   #FRK_JsonHeader := FALSE;
   #Line := WSTRING#'{';
   #Ok := "FRK_JsonAdd"(Key := 'set', Value := STRING_TO_WSTRING(#Data.SetName), Quoted := TRUE, LastField := FALSE, Line := #Line);
   IF NOT #Ok THEN
       #Line := WSTRING#'';
       RETURN;
   END_IF;
   #Ok := "FRK_JsonAdd"(Key := 'root', Value := STRING_TO_WSTRING(#Data.RootIdentity), Quoted := TRUE, LastField := FALSE, Line := #Line);
   IF NOT #Ok THEN
       #Line := WSTRING#'';
       RETURN;
   END_IF;
   #Ok := "FRK_JsonAdd"(Key := 'schema', Value := UINT_TO_WSTRING(#Data.SetSchema), Quoted := FALSE, LastField := FALSE, Line := #Line);
   IF NOT #Ok THEN
       #Line := WSTRING#'';
       RETURN;
   END_IF;
   #Ok := "FRK_JsonAdd"(Key := 'configRev', Value := UDINT_TO_WSTRING(#Data.ConfigRev), Quoted := FALSE, LastField := FALSE, Line := #Line);
   IF NOT #Ok THEN
       #Line := WSTRING#'';
       RETURN;
   END_IF;
   #Ok := "FRK_JsonAdd"(Key := 'kind', Value := DINT_TO_WSTRING(#Data.Kind), Quoted := FALSE, LastField := FALSE, Line := #Line);
   IF NOT #Ok THEN
       #Line := WSTRING#'';
       RETURN;
   END_IF;
   #Ok := "FRK_JsonAdd"(Key := 'model', Value := STRING_TO_WSTRING(#Data.ModelCode), Quoted := TRUE, LastField := FALSE, Line := #Line);
   IF NOT #Ok THEN
       #Line := WSTRING#'';
       RETURN;
   END_IF;
   #Ok := "FRK_JsonAdd"(Key := 'records', Value := DINT_TO_WSTRING(#Data.RecordCount), Quoted := FALSE, LastField := FALSE, Line := #Line);
   IF NOT #Ok THEN
       #Line := WSTRING#'';
       RETURN;
   END_IF;
   #Ok := "FRK_JsonAdd"(Key := 'created', Value := ULINT_TO_WSTRING(LDT_TO_ULINT(#Data.CreatedAt) / ULINT#1000000000), Quoted := FALSE, LastField := FALSE, Line := #Line);
   IF NOT #Ok THEN
       #Line := WSTRING#'';
       RETURN;
   END_IF;
   IF #Data.TimeSynchronized THEN
       #Flag := WSTRING#'1';
   ELSE
       #Flag := WSTRING#'0';
   END_IF;
   #Ok := "FRK_JsonAdd"(Key := 'clock', Value := #Flag, Quoted := FALSE, LastField := TRUE, Line := #Line);
   IF NOT #Ok THEN
       #Line := WSTRING#'';
       RETURN;
   END_IF;
   #FRK_JsonHeader := TRUE;
END_FUNCTION

FUNCTION "FRK_JsonParse" : Bool   // FC110, SCL
{ S7_Optimized_Access := 'TRUE' }
VERSION : 0.1
// Strict flat JSON object scanner: whole object, unique known fields, exact
//  types, numeric integer grammar; strings decode escapes before owner checks.
// stored: AutoNumber true, IsIECCheckEnabled false, SetENOAutomatically false, UDAEnableTagReadback false
   VAR_INPUT
      Line : WString;
   END_VAR
   VAR_IN_OUT
      Fields : Array[1..9] of "FRK_JsonField";
      Count : Int;
   END_VAR
   VAR_TEMP
      Pos : Int;
      Limit : Int;
      Digit : Int;
      CodePoint : UInt;
      HexIndex : Int;
      Index : Int;
      Part : Int;
      Text : WString[160];
      Piece : WString[1];
      Quoted : Bool;
      Closed : Bool;
      Ch : WChar;
   END_VAR
BEGIN

   #FRK_JsonParse := FALSE;
   #Count := 0;
   #Pos := 1;
   #Limit := LEN(#Line);
   IF #Limit < 2 OR #Line[#Pos] <> WCHAR#'{' THEN
       RETURN;
   END_IF;
   #Pos := #Pos + 1;
   WHILE #Pos <= #Limit DO
       "FRK_JsonSkip"(Line := #Line,
                      Pos := #Pos);
       IF #Pos > #Limit OR #Count >= 9 THEN
           RETURN;
       END_IF;
       #Count := #Count + 1;
       FOR #Part := 1 TO 2 DO
           #Text := WSTRING#'';
           #Closed := FALSE;
           #Quoted := #Line[#Pos] = WCHAR#'"';
           IF #Part = 1 AND NOT #Quoted THEN
               RETURN;
           END_IF;
           IF #Quoted THEN
               #Pos := #Pos + 1;
           END_IF;
           WHILE #Pos <= #Limit DO
               #Ch := #Line[#Pos];
               IF #Quoted AND #Ch = WCHAR#'"' THEN
                   #Closed := TRUE;
                   #Pos := #Pos + 1;
                   EXIT;
               END_IF;
               IF NOT #Quoted AND (#Ch = WCHAR#',' OR #Ch = WCHAR#'}' OR #Ch = WCHAR#' ') THEN
                   #Closed := TRUE;
                   EXIT;
               END_IF;
               IF #Ch < WCHAR#'$0020' THEN
                   RETURN;
               END_IF;
               IF #Quoted AND #Ch = WCHAR#'\' THEN
                   #Pos := #Pos + 1;
                   IF #Pos > #Limit THEN
                       RETURN;
                   END_IF;
                   #Ch := #Line[#Pos];
                   IF #Ch = WCHAR#'u' THEN
                       #CodePoint := 0;
                       FOR #HexIndex := 1 TO 4 DO
                           #Pos := #Pos + 1;
                           IF #Pos > #Limit THEN
                               RETURN;
                           END_IF;
                           #Ch := #Line[#Pos];
                           #Digit := -1;
                           IF #Ch >= WCHAR#'0' AND #Ch <= WCHAR#'9' THEN
                               #Digit := WORD_TO_INT(WCHAR_TO_WORD(#Ch)) - 48;
                           ELSIF #Ch >= WCHAR#'a' AND #Ch <= WCHAR#'f' THEN
                               #Digit := WORD_TO_INT(WCHAR_TO_WORD(#Ch)) - 87;
                           ELSIF #Ch >= WCHAR#'A' AND #Ch <= WCHAR#'F' THEN
                               #Digit := WORD_TO_INT(WCHAR_TO_WORD(#Ch)) - 55;
                           END_IF;
                           IF #Digit < 0 THEN
                               RETURN;
                           END_IF;
                           #CodePoint := #CodePoint * 16 + INT_TO_UINT(#Digit);
                       END_FOR;
                       IF #CodePoint = 0 OR #CodePoint >= UINT#16#D000 THEN
                           RETURN;
                       END_IF;
                       #Ch := WORD_TO_WCHAR(UINT_TO_WORD(#CodePoint));
                   ELSIF #Ch = WCHAR#'n' THEN
                       #Ch := WCHAR#'$000A';
                   ELSIF #Ch = WCHAR#'r' THEN
                       #Ch := WCHAR#'$000D';
                   ELSIF #Ch = WCHAR#'t' THEN
                       #Ch := WCHAR#'$0009';
                   ELSIF #Ch = WCHAR#'b' THEN
                       #Ch := WCHAR#'$0008';
                   ELSIF #Ch = WCHAR#'f' THEN
                       #Ch := WCHAR#'$000C';
                   ELSIF #Ch <> WCHAR#'"' AND #Ch <> WCHAR#'\' AND #Ch <> WCHAR#'/' THEN
                       RETURN;
                   END_IF;
               ELSIF NOT #Quoted AND (#Ch < WCHAR#'0' OR #Ch > WCHAR#'9') THEN
                   RETURN;
               END_IF;
               IF LEN(#Text) >= 160 THEN
                   RETURN;
               END_IF;
               #Piece := WSTRING#' ';
               #Piece[1] := #Ch;
               #Text := CONCAT(IN1 := #Text, IN2 := #Piece);
               #Pos := #Pos + 1;
           END_WHILE;
           IF NOT #Closed THEN
               RETURN;
           END_IF;
           IF #Part = 1 THEN
               IF LEN(#Text) < 1 OR LEN(#Text) > 16 THEN
                   RETURN;
               END_IF;
               #Fields[#Count].Key := WSTRING_TO_STRING(#Text);
               FOR #Index := 1 TO #Count - 1 DO
                   IF #Fields[#Index].Key = #Fields[#Count].Key THEN
                       RETURN;
                   END_IF;
               END_FOR;
               "FRK_JsonSkip"(Line := #Line,
                              Pos := #Pos);
               IF #Pos > #Limit THEN
                   RETURN;
               END_IF;
               IF #Line[#Pos] <> WCHAR#':' THEN
                   RETURN;
               END_IF;
               #Pos := #Pos + 1;
               "FRK_JsonSkip"(Line := #Line,
                              Pos := #Pos);
               IF #Pos > #Limit THEN
                   RETURN;
               END_IF;
           ELSE
               IF NOT #Quoted AND (LEN(#Text) = 0 OR (LEN(#Text) > 1 AND #Text[1] = WCHAR#'0')) THEN
                   RETURN;
               END_IF;
               #Fields[#Count].Text := #Text;
               #Fields[#Count].Quoted := #Quoted;
           END_IF;
       END_FOR;
       "FRK_JsonSkip"(Line := #Line,
                      Pos := #Pos);
       IF #Pos > #Limit THEN
           RETURN;
       END_IF;
       IF #Line[#Pos] = WCHAR#'}' THEN
           #Pos := #Pos + 1;
           "FRK_JsonSkip"(Line := #Line,
                          Pos := #Pos);
           #FRK_JsonParse := #Pos > #Limit;
           RETURN;
       END_IF;
       IF #Line[#Pos] <> WCHAR#',' THEN
           RETURN;
       END_IF;
       #Pos := #Pos + 1;
   END_WHILE;
END_FUNCTION

FUNCTION "FRK_JsonPut" : Bool   // FC108, SCL
{ S7_Optimized_Access := 'TRUE' }
VERSION : 0.1
// Append complete text or refuse. Explicit destination width and length check
//  protect long WSTRING lines against truncation in the Siemens string runtime.
// stored: AutoNumber true, IsIECCheckEnabled false, SetENOAutomatically false, UDAEnableTagReadback false
   VAR_INPUT
      Text : WString;
   END_VAR
   VAR_IN_OUT
      Line : WString;
   END_VAR
   VAR_TEMP
      Expected : Int;
   END_VAR
BEGIN

   #FRK_JsonPut := FALSE;
   #Expected := LEN(#Line) + LEN(#Text);
   IF #Expected > 480 THEN
       RETURN;
   END_IF;
   #Line := CONCAT(IN1 := #Line, IN2 := #Text);
   #FRK_JsonPut := LEN(#Line) = #Expected;
END_FUNCTION

FUNCTION "FRK_JsonReadHeader" : Bool   // FC119, SCL
{ S7_Optimized_Access := 'TRUE' }
VERSION : 0.1
// stored: AutoNumber true, IsIECCheckEnabled false, SetENOAutomatically false, UDAEnableTagReadback false
   VAR_INPUT
      Count : Int;
      Fields : Array[1..9] of "FRK_JsonField";
   END_VAR
   VAR_IN_OUT
      Data : "ST_ConfigSetInfo";
   END_VAR
   VAR_TEMP
      Candidate : "ST_ConfigSetInfo";
      Index : Int;
      Found : Int;
      Ok : Bool;
   END_VAR
BEGIN

   #FRK_JsonReadHeader := FALSE;
   IF #Count <> 9 THEN
       RETURN;
   END_IF;
   #Found := 0;
   FOR #Index := 1 TO #Count DO
       IF #Fields[#Index].Key = 'set' THEN
           #Found := #Index;
       END_IF;
   END_FOR;
   IF #Found = 0 THEN
       RETURN;
   END_IF;
   IF #Fields[#Found].Quoted <> TRUE THEN
       RETURN;
   END_IF;
   IF LEN(#Fields[#Found].Text) > 80 OR STRING_TO_WSTRING(WSTRING_TO_STRING(#Fields[#Found].Text)) <> #Fields[#Found].Text THEN
       RETURN;
   END_IF;
   #Candidate.SetName := WSTRING_TO_STRING(#Fields[#Found].Text);
   #Found := 0;
   FOR #Index := 1 TO #Count DO
       IF #Fields[#Index].Key = 'root' THEN
           #Found := #Index;
       END_IF;
   END_FOR;
   IF #Found = 0 THEN
       RETURN;
   END_IF;
   IF #Fields[#Found].Quoted <> TRUE THEN
       RETURN;
   END_IF;
   IF LEN(#Fields[#Found].Text) > 80 OR STRING_TO_WSTRING(WSTRING_TO_STRING(#Fields[#Found].Text)) <> #Fields[#Found].Text THEN
       RETURN;
   END_IF;
   #Candidate.RootIdentity := WSTRING_TO_STRING(#Fields[#Found].Text);
   #Found := 0;
   FOR #Index := 1 TO #Count DO
       IF #Fields[#Index].Key = 'schema' THEN
           #Found := #Index;
       END_IF;
   END_FOR;
   IF #Found = 0 THEN
       RETURN;
   END_IF;
   IF #Fields[#Found].Quoted <> FALSE THEN
       RETURN;
   END_IF;
   #Ok := "FRK_ConfigDecode"(Text := #Fields[#Found].Text, Storage := 4, Minimum := 0.0, Maximum := 65535.0, MaxLength := 0, Value := "FRK_ConfigScratch".Value);
   IF NOT #Ok THEN
       RETURN;
   END_IF;
   #Candidate.SetSchema := LINT_TO_UINT("FRK_ConfigScratch".Value.Number);
   #Found := 0;
   FOR #Index := 1 TO #Count DO
       IF #Fields[#Index].Key = 'configRev' THEN
           #Found := #Index;
       END_IF;
   END_FOR;
   IF #Found = 0 THEN
       RETURN;
   END_IF;
   IF #Fields[#Found].Quoted <> FALSE THEN
       RETURN;
   END_IF;
   #Ok := "FRK_ConfigDecode"(Text := #Fields[#Found].Text, Storage := 4, Minimum := 0.0, Maximum := 4294967295.0, MaxLength := 0, Value := "FRK_ConfigScratch".Value);
   IF NOT #Ok THEN
       RETURN;
   END_IF;
   #Candidate.ConfigRev := LINT_TO_UDINT("FRK_ConfigScratch".Value.Number);
   #Found := 0;
   FOR #Index := 1 TO #Count DO
       IF #Fields[#Index].Key = 'kind' THEN
           #Found := #Index;
       END_IF;
   END_FOR;
   IF #Found = 0 THEN
       RETURN;
   END_IF;
   IF #Fields[#Found].Quoted <> FALSE THEN
       RETURN;
   END_IF;
   #Ok := "FRK_ConfigDecode"(Text := #Fields[#Found].Text, Storage := 4, Minimum := 0.0, Maximum := 1.0, MaxLength := 0, Value := "FRK_ConfigScratch".Value);
   IF NOT #Ok THEN
       RETURN;
   END_IF;
   #Candidate.Kind := LINT_TO_DINT("FRK_ConfigScratch".Value.Number);
   #Found := 0;
   FOR #Index := 1 TO #Count DO
       IF #Fields[#Index].Key = 'model' THEN
           #Found := #Index;
       END_IF;
   END_FOR;
   IF #Found = 0 THEN
       RETURN;
   END_IF;
   IF #Fields[#Found].Quoted <> TRUE THEN
       RETURN;
   END_IF;
   IF LEN(#Fields[#Found].Text) > 64 OR STRING_TO_WSTRING(WSTRING_TO_STRING(#Fields[#Found].Text)) <> #Fields[#Found].Text THEN
       RETURN;
   END_IF;
   #Candidate.ModelCode := WSTRING_TO_STRING(#Fields[#Found].Text);
   #Found := 0;
   FOR #Index := 1 TO #Count DO
       IF #Fields[#Index].Key = 'records' THEN
           #Found := #Index;
       END_IF;
   END_FOR;
   IF #Found = 0 THEN
       RETURN;
   END_IF;
   IF #Fields[#Found].Quoted <> FALSE THEN
       RETURN;
   END_IF;
   #Ok := "FRK_ConfigDecode"(Text := #Fields[#Found].Text, Storage := 4, Minimum := 0.0, Maximum := 3.0, MaxLength := 0, Value := "FRK_ConfigScratch".Value);
   IF NOT #Ok THEN
       RETURN;
   END_IF;
   #Candidate.RecordCount := LINT_TO_INT("FRK_ConfigScratch".Value.Number);
   #Found := 0;
   FOR #Index := 1 TO #Count DO
       IF #Fields[#Index].Key = 'created' THEN
           #Found := #Index;
       END_IF;
   END_FOR;
   IF #Found = 0 THEN
       RETURN;
   END_IF;
   IF #Fields[#Found].Quoted <> FALSE THEN
       RETURN;
   END_IF;
   #Ok := "FRK_ConfigDecode"(Text := #Fields[#Found].Text, Storage := 4, Minimum := 0.0, Maximum := 4294967295.0, MaxLength := 0, Value := "FRK_ConfigScratch".Value);
   IF NOT #Ok THEN
       RETURN;
   END_IF;
   #Candidate.CreatedAt := ULINT_TO_LDT(LINT_TO_ULINT("FRK_ConfigScratch".Value.Number) * ULINT#1000000000);
   #Found := 0;
   FOR #Index := 1 TO #Count DO
       IF #Fields[#Index].Key = 'clock' THEN
           #Found := #Index;
       END_IF;
   END_FOR;
   IF #Found = 0 THEN
       RETURN;
   END_IF;
   IF #Fields[#Found].Quoted <> FALSE THEN
       RETURN;
   END_IF;
   #Ok := "FRK_ConfigDecode"(Text := #Fields[#Found].Text, Storage := 4, Minimum := 0.0, Maximum := 1.0, MaxLength := 0, Value := "FRK_ConfigScratch".Value);
   IF NOT #Ok THEN
       RETURN;
   END_IF;
   #Candidate.TimeSynchronized := "FRK_ConfigScratch".Value.Number = 1;
   #Data := #Candidate;
   #FRK_JsonReadHeader := TRUE;
END_FUNCTION

FUNCTION "FRK_JsonReadRecord" : Bool   // FC121, SCL
{ S7_Optimized_Access := 'TRUE' }
VERSION : 0.1
// stored: AutoNumber true, IsIECCheckEnabled false, SetENOAutomatically false, UDAEnableTagReadback false
   VAR_INPUT
      Count : Int;
      Fields : Array[1..9] of "FRK_JsonField";
   END_VAR
   VAR_IN_OUT
      Data : "ST_ConfigRecord";
   END_VAR
   VAR_TEMP
      Candidate : "ST_ConfigRecord";
      Index : Int;
      Found : Int;
      Ok : Bool;
   END_VAR
BEGIN

   #FRK_JsonReadRecord := FALSE;
   IF #Count <> 6 THEN
       RETURN;
   END_IF;
   #Found := 0;
   FOR #Index := 1 TO #Count DO
       IF #Fields[#Index].Key = 'scope' THEN
           #Found := #Index;
       END_IF;
   END_FOR;
   IF #Found = 0 THEN
       RETURN;
   END_IF;
   IF #Fields[#Found].Quoted <> TRUE THEN
       RETURN;
   END_IF;
   IF LEN(#Fields[#Found].Text) > 80 OR STRING_TO_WSTRING(WSTRING_TO_STRING(#Fields[#Found].Text)) <> #Fields[#Found].Text THEN
       RETURN;
   END_IF;
   #Candidate.Scope := WSTRING_TO_STRING(#Fields[#Found].Text);
   #Found := 0;
   FOR #Index := 1 TO #Count DO
       IF #Fields[#Index].Key = 'key' THEN
           #Found := #Index;
       END_IF;
   END_FOR;
   IF #Found = 0 THEN
       RETURN;
   END_IF;
   IF #Fields[#Found].Quoted <> TRUE THEN
       RETURN;
   END_IF;
   IF LEN(#Fields[#Found].Text) > 160 OR STRING_TO_WSTRING(WSTRING_TO_STRING(#Fields[#Found].Text)) <> #Fields[#Found].Text THEN
       RETURN;
   END_IF;
   #Candidate.WriteKey := WSTRING_TO_STRING(#Fields[#Found].Text);
   #Found := 0;
   FOR #Index := 1 TO #Count DO
       IF #Fields[#Index].Key = 'rev' THEN
           #Found := #Index;
       END_IF;
   END_FOR;
   IF #Found = 0 THEN
       RETURN;
   END_IF;
   IF #Fields[#Found].Quoted <> FALSE THEN
       RETURN;
   END_IF;
   #Ok := "FRK_ConfigDecode"(Text := #Fields[#Found].Text, Storage := 4, Minimum := 0.0, Maximum := 4294967295.0, MaxLength := 0, Value := "FRK_ConfigScratch".Value);
   IF NOT #Ok THEN
       RETURN;
   END_IF;
   #Candidate.Revision := LINT_TO_UDINT("FRK_ConfigScratch".Value.Number);
   #Found := 0;
   FOR #Index := 1 TO #Count DO
       IF #Fields[#Index].Key = 'kind' THEN
           #Found := #Index;
       END_IF;
   END_FOR;
   IF #Found = 0 THEN
       RETURN;
   END_IF;
   IF #Fields[#Found].Quoted <> FALSE THEN
       RETURN;
   END_IF;
   #Ok := "FRK_ConfigDecode"(Text := #Fields[#Found].Text, Storage := 4, Minimum := 0.0, Maximum := 1.0, MaxLength := 0, Value := "FRK_ConfigScratch".Value);
   IF NOT #Ok THEN
       RETURN;
   END_IF;
   #Candidate.Kind := LINT_TO_DINT("FRK_ConfigScratch".Value.Number);
   #Found := 0;
   FOR #Index := 1 TO #Count DO
       IF #Fields[#Index].Key = 'type' THEN
           #Found := #Index;
       END_IF;
   END_FOR;
   IF #Found = 0 THEN
       RETURN;
   END_IF;
   IF #Fields[#Found].Quoted <> FALSE THEN
       RETURN;
   END_IF;
   #Ok := "FRK_ConfigDecode"(Text := #Fields[#Found].Text, Storage := 4, Minimum := 0.0, Maximum := 3.0, MaxLength := 0, Value := "FRK_ConfigScratch".Value);
   IF NOT #Ok THEN
       RETURN;
   END_IF;
   #Candidate.ValueType := LINT_TO_DINT("FRK_ConfigScratch".Value.Number);
   #Found := 0;
   FOR #Index := 1 TO #Count DO
       IF #Fields[#Index].Key = 'value' THEN
           #Found := #Index;
       END_IF;
   END_FOR;
   IF #Found = 0 THEN
       RETURN;
   END_IF;
   IF #Fields[#Found].Quoted <> TRUE THEN
       RETURN;
   END_IF;
   IF LEN(#Fields[#Found].Text) > 80 OR STRING_TO_WSTRING(WSTRING_TO_STRING(#Fields[#Found].Text)) <> #Fields[#Found].Text THEN
       RETURN;
   END_IF;
   #Candidate.ValueText := WSTRING_TO_STRING(#Fields[#Found].Text);
   #Data := #Candidate;
   #FRK_JsonReadRecord := TRUE;
END_FUNCTION

FUNCTION "FRK_JsonRecord" : Bool   // FC120, SCL
{ S7_Optimized_Access := 'TRUE' }
VERSION : 0.1
// stored: AutoNumber true, IsIECCheckEnabled false, SetENOAutomatically false, UDAEnableTagReadback false
   VAR_INPUT
      Data : "ST_ConfigRecord";
   END_VAR
   VAR_IN_OUT
      Line : WString;
   END_VAR
   VAR_TEMP
      Ok : Bool;
      Flag : WString[1];
   END_VAR
BEGIN

   #FRK_JsonRecord := FALSE;
   #Line := WSTRING#'{';
   #Ok := "FRK_JsonAdd"(Key := 'scope', Value := STRING_TO_WSTRING(#Data.Scope), Quoted := TRUE, LastField := FALSE, Line := #Line);
   IF NOT #Ok THEN
       #Line := WSTRING#'';
       RETURN;
   END_IF;
   #Ok := "FRK_JsonAdd"(Key := 'key', Value := STRING_TO_WSTRING(#Data.WriteKey), Quoted := TRUE, LastField := FALSE, Line := #Line);
   IF NOT #Ok THEN
       #Line := WSTRING#'';
       RETURN;
   END_IF;
   #Ok := "FRK_JsonAdd"(Key := 'rev', Value := UDINT_TO_WSTRING(#Data.Revision), Quoted := FALSE, LastField := FALSE, Line := #Line);
   IF NOT #Ok THEN
       #Line := WSTRING#'';
       RETURN;
   END_IF;
   #Ok := "FRK_JsonAdd"(Key := 'kind', Value := DINT_TO_WSTRING(#Data.Kind), Quoted := FALSE, LastField := FALSE, Line := #Line);
   IF NOT #Ok THEN
       #Line := WSTRING#'';
       RETURN;
   END_IF;
   #Ok := "FRK_JsonAdd"(Key := 'type', Value := DINT_TO_WSTRING(#Data.ValueType), Quoted := FALSE, LastField := FALSE, Line := #Line);
   IF NOT #Ok THEN
       #Line := WSTRING#'';
       RETURN;
   END_IF;
   #Ok := "FRK_JsonAdd"(Key := 'value', Value := STRING_TO_WSTRING(#Data.ValueText), Quoted := TRUE, LastField := TRUE, Line := #Line);
   IF NOT #Ok THEN
       #Line := WSTRING#'';
       RETURN;
   END_IF;
   #FRK_JsonRecord := TRUE;
END_FUNCTION

FUNCTION "FRK_JsonSkip" : Void   // FC113, SCL
{ S7_Optimized_Access := 'TRUE' }
VERSION : 0.1
// stored: AutoNumber true, IsIECCheckEnabled false, SetENOAutomatically false, UDAEnableTagReadback false
   VAR_INPUT
      Line : WString;
   END_VAR
   VAR_IN_OUT
      Pos : Int;
   END_VAR
BEGIN

   WHILE #Pos <= LEN(#Line) DO
       IF #Line[#Pos] <> WCHAR#' ' AND #Line[#Pos] <> WCHAR#'$0009' AND #Line[#Pos] <> WCHAR#'$000A' AND #Line[#Pos] <> WCHAR#'$000D' THEN
           RETURN;
       END_IF;
       #Pos := #Pos + 1;
   END_WHILE;
END_FUNCTION

FUNCTION "FRK_ManualApply" : Void   // FC82, SCL
{ S7_Optimized_Access := 'TRUE' }
VERSION : 0.1
// stored: AutoNumber true, IsIECCheckEnabled false, SetENOAutomatically false, UDAEnableTagReadback false
   VAR_INPUT
      Request : "ST_HmiRequest";
      Status : "ST_ModuleStatus";
      Core : "FRK_Core";
      Commands : Array[1..12] of "ST_CommandInfo";
      Count : DInt;
      Conditions : Array[1..16] of "FRK_ManualConditionRow";
   END_VAR
   VAR_IN_OUT
      Report : "ST_ReleaseReport";
      Execute : Bool;
      Command : DInt;
      ManualOwned : Bool;
   END_VAR
   VAR_TEMP
      Index : Int;
      Supported : Bool;
      PreviousCount : Int;
   END_VAR
BEGIN

   #Supported := FALSE;
   IF #Count >= 0 AND #Count <= 12 THEN
       FOR #Index := 1 TO DINT_TO_INT(#Count) DO
           IF #Commands[#Index].Value = #Request.IntValue AND #Commands[#Index].Style = 0 THEN
               #Supported := TRUE;
           END_IF;
       END_FOR;
   END_IF;
   IF NOT #Supported THEN
       "FRK_ReleaseReason"(Report := #Report,
                           Description := WSTRING#'std.error.unsupportedHmiRequest',
                           Reason := 2008,
                           Path := STRING_TO_WSTRING(#Status.Name),
                           Kind := 4);
   END_IF;
   IF #Core.Exec <> 0 OR #Execute OR #Core.ReleasePending THEN
       "FRK_ReleaseReason"(Report := #Report,
                           Description := WSTRING#'std.error.hmiRequestRejected',
                           Reason := 2011,
                           Path := STRING_TO_WSTRING(#Status.Name),
                           Kind := 4);
   END_IF;
   FOR #Index := 1 TO 16 DO
       IF #Conditions[#Index].Used AND NOT #Conditions[#Index].Ok THEN
           IF #Conditions[#Index].Value = 0 OR #Conditions[#Index].Value = #Request.IntValue THEN
               #PreviousCount := #Report.Count;
               "FRK_ReleaseReason"(Report := #Report,
                                   Description := #Conditions[#Index].Diag.Description,
                                   Reason := #Conditions[#Index].Diag.ReasonCode,
                                   Path := STRING_TO_WSTRING(#Status.Name),
                                   Kind := 3);
               IF #Report.Count > #PreviousCount THEN
                   #Report.Reasons[#Report.Count].Bypassable := #Conditions[#Index].Bypassable;
               END_IF;
           END_IF;
       END_IF;
   END_FOR;
   IF #Request.Kind = 11 AND #Report.Released THEN
       #Command := #Request.IntValue;
       #Execute := TRUE;
       #ManualOwned := TRUE;
   END_IF;
END_FUNCTION

FUNCTION "FRK_ManualCommon" : Void   // FC80, SCL
{ S7_Optimized_Access := 'TRUE' }
VERSION : 0.1
// stored: AutoNumber true, IsIECCheckEnabled false, SetENOAutomatically false, UDAEnableTagReadback false
   VAR_INPUT
      Core : "FRK_Core";
      Unit : "FRK_Unit";
      Status : "ST_ModuleStatus";
   END_VAR
   VAR_IN_OUT
      Report : "ST_ReleaseReport";
   END_VAR
BEGIN

   IF #Unit.Mode <> 1 OR #Unit.ModePending THEN
       "FRK_ReleaseReason"(Report := #Report,
                           Description := WSTRING#'std.release.manualModeRequired',
                           Reason := 2002,
                           Path := STRING_TO_WSTRING(#Status.Name),
                           Kind := 0);
   END_IF;
   IF #Core.Exec <> 0 OR #Unit.Clearing OR #Unit.FaultLatched THEN
       "FRK_ReleaseReason"(Report := #Report,
                           Description := WSTRING#'std.error.hmiRequestRejected',
                           Reason := 2011,
                           Path := STRING_TO_WSTRING(#Status.Name),
                           Kind := 4);
   END_IF;
   IF #Unit.AlarmBlocking THEN
       "FRK_ReleaseReason"(Report := #Report,
                           Description := WSTRING#'std.release.manualReset',
                           Reason := 0,
                           Path := STRING_TO_WSTRING(#Status.Name),
                           Kind := 2);
   END_IF;
   IF NOT #Unit.Permit THEN
       "FRK_ReleaseReason"(Report := #Report,
                           Description := #Unit.PermitDiag.Description,
                           Reason := #Unit.PermitDiag.ReasonCode,
                           Path := #Unit.PermitDiag.SourcePath,
                           Kind := 3);
   END_IF;
END_FUNCTION

FUNCTION "FRK_ManualCondition" : Void   // FC81, SCL
{ S7_Optimized_Access := 'TRUE' }
VERSION : 0.1
// stored: AutoNumber true, IsIECCheckEnabled false, SetENOAutomatically false, UDAEnableTagReadback false
   VAR_INPUT
      Slot : Int;
      Value : DInt;
      Ok : Bool;
      Diag : "ST_Diagnostic";
      Bypassable : Bool;
   END_VAR
   VAR_IN_OUT
      Conditions : Array[1..16] of "FRK_ManualConditionRow";
   END_VAR
BEGIN

   IF #Slot < 1 OR #Slot > 16 THEN
       RETURN;
   END_IF;
   #Conditions[#Slot].Used := TRUE;
   #Conditions[#Slot].Value := #Value;
   #Conditions[#Slot].Ok := #Ok;
   #Conditions[#Slot].Diag := #Diag;
   #Conditions[#Slot].Bypassable := #Bypassable;
END_FUNCTION

FUNCTION "FRK_ManualFinish" : Void   // FC83, SCL
{ S7_Optimized_Access := 'TRUE' }
VERSION : 0.1
// stored: AutoNumber true, IsIECCheckEnabled false, SetENOAutomatically false, UDAEnableTagReadback false
   VAR_INPUT
      Core : "FRK_Core";
   END_VAR
   VAR_IN_OUT
      Execute : Bool;
      ManualOwned : Bool;
   END_VAR
BEGIN

   IF #ManualOwned AND #Core.Exec <> 1 THEN
       #Execute := FALSE;
       #ManualOwned := FALSE;
   END_IF;
END_FUNCTION

FUNCTION "FRK_PartAborted" : Void   // FC67, SCL
{ S7_Optimized_Access := 'TRUE' }
VERSION : 0.1
// stored: AutoNumber true, IsIECCheckEnabled false, SetENOAutomatically false, UDAEnableTagReadback false
   VAR_IN_OUT
      Core : "FRK_Core";
      Unit : "FRK_Unit";
      Status : "ST_ModuleStatus";
      Part : "ST_PartContext";
      AlarmLog : "FRK_AlarmLog";
   END_VAR
BEGIN

   IF #Unit.CarrierIndex = 0 OR NOT #Part.Present THEN
       RETURN;
   END_IF;
   #Part.Result.Verdict := 0;
   IF #Core.Exec = 3 AND #Part.Result.ReasonCode = 0 THEN
       #Part.Result.ReasonCode := #Status.Diagnostic.ReasonCode;
   END_IF;
   "FRK_PartEvent"(AlarmLog := #AlarmLog,
                   Reason := 2027,
                   Uid := #Part.Uid,
                   SourcePath := #Status.Name);
   #Part.Present := FALSE;
END_FUNCTION

FUNCTION "FRK_PartEvent" : Void   // FC63, SCL
{ S7_Optimized_Access := 'TRUE' }
VERSION : 0.1
// stored: AutoNumber true, IsIECCheckEnabled false, SetENOAutomatically false, UDAEnableTagReadback false
   VAR_INPUT
      Reason : DInt;
      Uid : String;
      SourcePath : String;
   END_VAR
   VAR_IN_OUT
      AlarmLog : "FRK_AlarmLog";
   END_VAR
   VAR_TEMP
      Description : WString[255];
   END_VAR
BEGIN

   CASE #Reason OF
       2024:
           #Description := WSTRING#'std.event.partReceived: ';
       2025:
           #Description := WSTRING#'std.event.partProcessingStarted: ';
       2026:
           #Description := WSTRING#'std.event.partProcessed: ';
       2027:
           #Description := WSTRING#'std.event.partAborted: ';
       ELSE
           #Description := WSTRING#'';
   END_CASE;
   #Description := CONCAT(IN1 := #Description, IN2 := STRING_TO_WSTRING(#Uid));
   "FRK_AlarmMessage"(AlarmLog := #AlarmLog,
                      Reason := #Reason,
                      Description := #Description,
                      SourcePath := STRING_TO_WSTRING(#SourcePath));
END_FUNCTION

FUNCTION "FRK_PartProcessed" : Bool   // FC66, SCL
{ S7_Optimized_Access := 'TRUE' }
VERSION : 0.1
// stored: AutoNumber true, IsIECCheckEnabled false, SetENOAutomatically false, UDAEnableTagReadback false
   VAR_INPUT
      Verdict : DInt;
      Reason : DInt;
   END_VAR
   VAR_IN_OUT
      Core : "FRK_Core";
      Unit : "FRK_Unit";
      Status : "ST_ModuleStatus";
      Part : "ST_PartContext";
      AlarmLog : "FRK_AlarmLog";
   END_VAR
   VAR_TEMP
      Index : DInt;
      Stamp : DTL;
      ResultCode : Int;
   END_VAR
BEGIN

   #FRK_PartProcessed := FALSE;
   #Index := #Unit.CarrierIndex;
   IF #Index = 0 OR NOT #Part.Present THEN
       RETURN;
   END_IF;
   IF #Verdict < 1 OR #Verdict > 3 OR (#Verdict = 2 AND #Reason = 0) THEN
       "FRK_Fault"(Core := #Core,
                   Status := #Status,
                   ReasonCode := 2023,
                   Description := WSTRING#'std.error.nokReasonRequired');
       RETURN;
   END_IF;
   IF #Index < 1 OR #Index > 4 THEN
       "FRK_Fault"(Core := #Core,
                   Status := #Status,
                   ReasonCode := 2021,
                   Description := WSTRING#'std.error.partCarrierWriteFailed');
       RETURN;
   END_IF;
   IF NOT "FRK_Carriers".Slots[#Index].Enabled THEN
       "FRK_Fault"(Core := #Core,
                   Status := #Status,
                   ReasonCode := 2021,
                   Description := WSTRING#'std.error.partCarrierWriteFailed');
       RETURN;
   END_IF;
   IF #Part.Uid <> "FRK_Carriers".Slots[#Index].Context.Uid THEN
       "FRK_Fault"(Core := #Core,
                   Status := #Status,
                   ReasonCode := 2022,
                   Description := WSTRING#'std.error.partCarrierReadFailed');
       RETURN;
   END_IF;
   #Part.Result.Verdict := #Verdict;
   #Part.Result.ReasonCode := #Reason;
   #Part.Result.StationPath := STRING_TO_WSTRING(#Status.Name);
   #Part.Result.TimeSynchronized := FALSE;
   #ResultCode := RD_SYS_T(OUT => #Stamp);
   IF #ResultCode = 0 THEN
       #Part.Result.Stamp := DTL_TO_LDT(#Stamp);
   END_IF;
   "FRK_Carriers".Slots[#Index].Written := #Part;
   IF "FRK_Carriers".Slots[#Index].Writes < UDINT#4294967295 THEN
       "FRK_Carriers".Slots[#Index].Writes := "FRK_Carriers".Slots[#Index].Writes + 1;
   END_IF;
   CASE #Verdict OF
       1:
           IF #Unit.Good < UDINT#4294967295 THEN
               #Unit.Good := #Unit.Good + 1;
           END_IF;
       2:
           IF #Unit.Nok < UDINT#4294967295 THEN
               #Unit.Nok := #Unit.Nok + 1;
           END_IF;
           #Unit.NokReason := #Reason;
       3:
           IF #Unit.Rework < UDINT#4294967295 THEN
               #Unit.Rework := #Unit.Rework + 1;
           END_IF;
       ELSE
           RETURN;
   END_CASE;
   // The provider result is written before publishing EVENT_PART_PROCESSED.
   "FRK_PartEvent"(AlarmLog := #AlarmLog,
                   Reason := 2026,
                   Uid := #Part.Uid,
                   SourcePath := #Status.Name);
   #Part.Present := FALSE;
   #FRK_PartProcessed := TRUE;
END_FUNCTION

FUNCTION "FRK_PartReceived" : Bool   // FC64, SCL
{ S7_Optimized_Access := 'TRUE' }
VERSION : 0.1
// stored: AutoNumber true, IsIECCheckEnabled false, SetENOAutomatically false, UDAEnableTagReadback false
   VAR_IN_OUT
      Core : "FRK_Core";
      Unit : "FRK_Unit";
      Status : "ST_ModuleStatus";
      Part : "ST_PartContext";
      AlarmLog : "FRK_AlarmLog";
   END_VAR
   VAR_TEMP
      Index : DInt;
      Uid : String[64];
      ResultIndex : DInt;
   END_VAR
BEGIN

   #FRK_PartReceived := FALSE;
   #Index := #Unit.CarrierIndex;
   IF #Index = 0 THEN
       RETURN;
   END_IF;
   IF #Index < 1 OR #Index > 4 THEN
       "FRK_Fault"(Core := #Core,
                   Status := #Status,
                   ReasonCode := 2020,
                   Description := WSTRING#'std.error.partCarrierReadFailed');
       RETURN;
   END_IF;
   IF NOT "FRK_Carriers".Slots[#Index].Enabled OR "FRK_Carriers".Slots[#Index].Kind <> 2 OR "FRK_Carriers".Slots[#Index].Serial = UDINT#4294967295 THEN
       "FRK_Fault"(Core := #Core,
                   Status := #Status,
                   ReasonCode := 2020,
                   Description := WSTRING#'std.error.partCarrierReadFailed');
       RETURN;
   END_IF;
   "FRK_Carriers".Slots[#Index].Serial := "FRK_Carriers".Slots[#Index].Serial + 1;
   #Uid := CONCAT(IN1 := 'FRK-', IN2 := DINT_TO_STRING(#Index));
   #Uid := CONCAT(IN1 := #Uid, IN2 := '-');
   #Uid := CONCAT(IN1 := #Uid, IN2 := UDINT_TO_STRING("FRK_Carriers".Slots[#Index].Serial));
   #Part.Uid := #Uid;
   #Part.Present := TRUE;
   #Part.CarrierKind := 2;
   #Part.Result.Verdict := 0;
   #Part.Result.ReasonCode := 0;
   #Part.Result.StationPath := STRING_TO_WSTRING(#Status.Name);
   #Part.Result.Stamp := LDT#1970-01-01-00:00:00.000000000;
   #Part.Result.TimeSynchronized := FALSE;
   FOR #ResultIndex := 1 TO 32 DO
       #Part.Result.Records[#ResultIndex].Name := '';
   END_FOR;
   FOR #ResultIndex := 1 TO 8 DO
       #Part.Parents[#ResultIndex] := '';
   END_FOR;
   "FRK_Carriers".Slots[#Index].Context := #Part;
   "FRK_PartEvent"(AlarmLog := #AlarmLog,
                   Reason := 2024,
                   Uid := #Part.Uid,
                   SourcePath := #Status.Name);
   #FRK_PartReceived := TRUE;
END_FUNCTION

FUNCTION "FRK_PartRecord" : Bool   // FC145, SCL
{ S7_Optimized_Access := 'TRUE' }
VERSION : 0.1
// stored: AutoNumber true, IsIECCheckEnabled false, SetENOAutomatically false, UDAEnableTagReadback false
   VAR_INPUT
      RecordName : String;
      Value : LReal;
      Minimum : LReal;
      Maximum : LReal;
      Target : LReal;
      EngUnit : String;
   END_VAR
   VAR_IN_OUT
      Core : "FRK_Core";
      Status : "ST_ModuleStatus";
      Part : "ST_PartContext";
   END_VAR
   VAR_TEMP
      Index : Int;
   END_VAR
BEGIN

   #FRK_PartRecord := FALSE;
   IF NOT #Part.Present THEN
       RETURN;
   END_IF;
   IF #RecordName = '' OR LEN(#RecordName) > 64 OR LEN(#EngUnit) > 16
       OR #Minimum > #Maximum OR #Value <> #Value OR #Minimum <> #Minimum OR #Maximum <> #Maximum OR #Target <> #Target THEN
       "FRK_Fault"(Core := #Core,
                   Status := #Status,
                   ReasonCode := 2023,
                   Description := WSTRING#'std.error.partRecordRejected');
       RETURN;
   END_IF;
   FOR #Index := 1 TO 32 DO
       IF #Part.Result.Records[#Index].Name = #RecordName OR #Part.Result.Records[#Index].Name = '' THEN
           #Part.Result.Records[#Index].Name := #RecordName;
           #Part.Result.Records[#Index].Value := #Value;
           #Part.Result.Records[#Index].Minimum := #Minimum;
           #Part.Result.Records[#Index].Maximum := #Maximum;
           #Part.Result.Records[#Index].Target := #Target;
           #Part.Result.Records[#Index].Unit := #EngUnit;
           #Part.Result.Records[#Index].InTol := #Value >= #Minimum AND #Value <= #Maximum;
           #FRK_PartRecord := TRUE;
           RETURN;
       END_IF;
   END_FOR;
   "FRK_Fault"(Core := #Core,
               Status := #Status,
               ReasonCode := 2023,
               Description := WSTRING#'std.error.partRecordTableFull');
END_FUNCTION

FUNCTION "FRK_PartStarted" : Void   // FC65, SCL
{ S7_Optimized_Access := 'TRUE' }
VERSION : 0.1
// stored: AutoNumber true, IsIECCheckEnabled false, SetENOAutomatically false, UDAEnableTagReadback false
   VAR_IN_OUT
      Unit : "FRK_Unit";
      Status : "ST_ModuleStatus";
      Part : "ST_PartContext";
      AlarmLog : "FRK_AlarmLog";
   END_VAR
BEGIN

   IF #Unit.CarrierIndex = 0 OR NOT #Part.Present THEN
       RETURN;
   END_IF;
   "FRK_PartEvent"(AlarmLog := #AlarmLog,
                   Reason := 2025,
                   Uid := #Part.Uid,
                   SourcePath := #Status.Name);
END_FUNCTION

FUNCTION "FRK_PathOwned" : Bool   // FC78, SCL
{ S7_Optimized_Access := 'TRUE' }
VERSION : 0.1
// Shared Unit routing: typed generated edges carry these owning predicates.
// stored: AutoNumber true, IsIECCheckEnabled false, SetENOAutomatically false, UDAEnableTagReadback false
   VAR_INPUT
      OwnerPath : String;
      TargetPath : WString;
   END_VAR
   VAR_TEMP
      Width : Int;
   END_VAR
BEGIN

   #FRK_PathOwned := FALSE;
   #Width := LEN(#OwnerPath);
   IF #Width = 0 THEN
       RETURN;
   END_IF;
   IF #TargetPath = STRING_TO_WSTRING(#OwnerPath) THEN
       #FRK_PathOwned := TRUE;
       RETURN;
   END_IF;
   IF LEN(#TargetPath) <= #Width THEN
       RETURN;
   END_IF;
   #FRK_PathOwned := LEFT(IN := #TargetPath, L := #Width) = STRING_TO_WSTRING(#OwnerPath) AND #TargetPath[#Width + 1] = WCHAR#'.';
END_FUNCTION

FUNCTION "FRK_Pending" : Void   // FC12, SCL
{ S7_Optimized_Access := 'TRUE' }
VERSION : 0.1
// stored: AutoNumber true, IsIECCheckEnabled false, SetENOAutomatically false, UDAEnableTagReadback false
   VAR_INPUT
      Diag : "ST_Diagnostic";
   END_VAR
   VAR_IN_OUT
      Core : "FRK_Core";
      Status : "ST_ModuleStatus";
   END_VAR
BEGIN

   IF #Core.Exec = 1 AND NOT #Core.DiagTouched THEN
       #Status.Diagnostic := #Diag;
       #Status.Diagnostic.Severity := 0;
       #Core.DiagTouched := TRUE;
   END_IF;
END_FUNCTION

FUNCTION "FRK_Rationalize" : Void   // FC6, SCL
{ S7_Optimized_Access := 'TRUE' }
VERSION : 0.1
// stored: AutoNumber true, IsIECCheckEnabled false, SetENOAutomatically false, UDAEnableTagReadback false
   VAR_IN_OUT
      Diag : "ST_Diagnostic";
   END_VAR
BEGIN

   CASE #Diag.ReasonCode OF
       10:
           #Diag.Severity := 1;
           #Diag.Category := 2;
       11:
           #Diag.Severity := 0;
           #Diag.Category := 2;
       12:
           #Diag.Severity := 0;
           #Diag.Category := 2;
       13:
           #Diag.Severity := 1;
           #Diag.Category := 2;
       14:
           #Diag.Severity := 1;
           #Diag.Category := 2;
       15:
           #Diag.Severity := 2;
           #Diag.Category := 2;
       16:
           #Diag.Severity := 0;
           #Diag.Category := 2;
       17:
           #Diag.Severity := 0;
           #Diag.Category := 2;
       18:
           #Diag.Severity := 1;
           #Diag.Category := 2;
       19:
           #Diag.Severity := 0;
           #Diag.Category := 2;
       20:
           #Diag.Severity := 1;
           #Diag.Category := 2;
       21:
           #Diag.Severity := 0;
           #Diag.Category := 2;
       2001:
           #Diag.Severity := 1;
           #Diag.Category := 0;
       2002:
           #Diag.Severity := 0;
           #Diag.Category := 0;
       2003:
           #Diag.Severity := 1;
           #Diag.Category := 0;
       2004:
           #Diag.Severity := 1;
           #Diag.Category := 0;
       2005:
           #Diag.Severity := 0;
           #Diag.Category := 0;
       2006:
           #Diag.Severity := 1;
           #Diag.Category := 0;
       2007:
           #Diag.Severity := 0;
           #Diag.Category := 0;
       2008:
           #Diag.Severity := 0;
           #Diag.Category := 0;
       2010:
           #Diag.Severity := 1;
           #Diag.Category := 2;
       2011:
           #Diag.Severity := 0;
           #Diag.Category := 0;
       2012:
           #Diag.Severity := 1;
           #Diag.Category := 2;
       2020:
           #Diag.Severity := 1;
           #Diag.Category := 2;
       2021:
           #Diag.Severity := 1;
           #Diag.Category := 2;
       2022:
           #Diag.Severity := 2;
           #Diag.Category := 0;
       2023:
           #Diag.Severity := 1;
           #Diag.Category := 0;
       2024:
           #Diag.Severity := 0;
           #Diag.Category := 0;
       2025:
           #Diag.Severity := 0;
           #Diag.Category := 0;
       2026:
           #Diag.Severity := 0;
           #Diag.Category := 0;
       2027:
           #Diag.Severity := 0;
           #Diag.Category := 0;
       2030:
           #Diag.Severity := 0;
           #Diag.Category := 2;
       2040:
           #Diag.Severity := 1;
           #Diag.Category := 2;
       2041:
           #Diag.Severity := 1;
           #Diag.Category := 2;
       2042:
           #Diag.Severity := 0;
           #Diag.Category := 2;
       2043:
           #Diag.Severity := 0;
           #Diag.Category := 2;
       2901:
           #Diag.Severity := 0;
           #Diag.Category := 2;
       ELSE
           RETURN;
   END_CASE;
END_FUNCTION

FUNCTION "FRK_RecordTiming" : Void   // FC17, SCL
{ S7_Optimized_Access := 'TRUE' }
VERSION : 0.1
// stored: AutoNumber true, IsIECCheckEnabled false, SetENOAutomatically false, UDAEnableTagReadback false
   VAR_IN_OUT
      Core : "FRK_Core";
   END_VAR
   VAR_TEMP
      Index : DInt;
      Slot : DInt;
      DurationMs : UDInt;
      AverageMs : LInt;
   END_VAR
BEGIN

   #DurationMs := "FRK_Elapsed"(NewMs := "FRK_Clock".NowMs, OldMs := #Core.StartMs);
   // TIME's positive domain is bounded; clamp instead of publishing negatives.
   IF #DurationMs > UDINT#2147483647 THEN
       #DurationMs := UDINT#2147483647;
   END_IF;
   #Core.Timing.LastCmdTime := DINT_TO_TIME(UDINT_TO_DINT(#DurationMs));
   #Slot := 0;
   FOR #Index := 1 TO 8 DO
       IF #Core.Timing.Rows[#Index].Count > 0 AND #Core.Timing.Rows[#Index].Id = #Core.Command THEN
           #Slot := #Index;
           EXIT;
       ELSIF #Slot = 0 AND #Core.Timing.Rows[#Index].Count = 0 THEN
           #Slot := #Index;
       END_IF;
   END_FOR;
   IF #Slot = 0 THEN
       #Core.Timing.Truncated := TRUE;
   ELSE
       #Core.Timing.Rows[#Slot].Id := #Core.Command;
       #Core.Timing.Rows[#Slot].Label := #Core.CommandLabel;
       IF #Core.Timing.Rows[#Slot].Count < UDINT#4294967295 THEN
           #Core.Timing.Rows[#Slot].Count := #Core.Timing.Rows[#Slot].Count + 1;
       END_IF;
       #Core.Timing.Rows[#Slot].Last := #Core.Timing.LastCmdTime;
       IF #Core.Timing.Rows[#Slot].Count = 1 OR #Core.Timing.LastCmdTime < #Core.Timing.Rows[#Slot].Minimum THEN
           #Core.Timing.Rows[#Slot].Minimum := #Core.Timing.LastCmdTime;
       END_IF;
       IF #Core.Timing.LastCmdTime > #Core.Timing.Rows[#Slot].Maximum THEN
           #Core.Timing.Rows[#Slot].Maximum := #Core.Timing.LastCmdTime;
       END_IF;
       #AverageMs := DINT_TO_LINT(TIME_TO_DINT(#Core.Timing.Rows[#Slot].Avg));
       #AverageMs := #AverageMs + (UDINT_TO_LINT(#DurationMs) - #AverageMs) / UDINT_TO_LINT(#Core.Timing.Rows[#Slot].Count);
       #Core.Timing.Rows[#Slot].Avg := DINT_TO_TIME(LINT_TO_DINT(#AverageMs));
   END_IF;
   #Core.TimingOpen := FALSE;
END_FUNCTION

FUNCTION "FRK_ReleaseCommand" : Void   // FC19, SCL
{ S7_Optimized_Access := 'TRUE' }
VERSION : 0.1
// stored: AutoNumber true, IsIECCheckEnabled false, SetENOAutomatically false, UDAEnableTagReadback false
   VAR_IN_OUT
      Core : "FRK_Core";
      Execute : Bool;
   END_VAR
BEGIN

   #Execute := FALSE;
   #Core.ReleasePending := TRUE;
END_FUNCTION

FUNCTION "FRK_ReleaseReason" : Void   // FC69, SCL
{ S7_Optimized_Access := 'TRUE' }
VERSION : 0.1
// stored: AutoNumber true, IsIECCheckEnabled false, SetENOAutomatically false, UDAEnableTagReadback false
   VAR_INPUT
      Description : WString;
      Reason : DInt;
      Path : WString;
      Kind : DInt;
   END_VAR
   VAR_IN_OUT
      Report : "ST_ReleaseReport";
   END_VAR
BEGIN

   #Report.Released := FALSE;
   IF #Report.Count < 24 THEN
       #Report.Count := #Report.Count + 1;
       #Report.Reasons[#Report.Count].Description := #Description;
       #Report.Reasons[#Report.Count].ReasonCode := #Reason;
       #Report.Reasons[#Report.Count].SourcePath := #Path;
       #Report.Reasons[#Report.Count].Kind := #Kind;
       #Report.Reasons[#Report.Count].Bypassable := FALSE;
   END_IF;
END_FUNCTION

FUNCTION "FRK_Release_PressDemoUnit" : Void   // FC171, SCL
{ S7_Optimized_Access := 'TRUE' }
VERSION : 0.1
// stored: AutoNumber true, IsIECCheckEnabled false, SetENOAutomatically false, UDAEnableTagReadback false
   VAR_IN_OUT
      Unit : "FRK_Unit";
      Hal : "ST_PressDemoUnitHal";
   END_VAR
BEGIN

   "FRK_UnitSetPermit"(Unit := #Unit,
                       Ok := #Hal.Process.AirPressureOk,
                       Diag := #Hal.Process.PermitDiagnostic);
END_FUNCTION

FUNCTION "FRK_RouteAbort" : Void   // FC16, SCL
{ S7_Optimized_Access := 'TRUE' }
VERSION : 0.1
// stored: AutoNumber true, IsIECCheckEnabled false, SetENOAutomatically false, UDAEnableTagReadback false
   VAR_INPUT
      Abort : Bool;
   END_VAR
   VAR_IN_OUT
      Core : "FRK_Core";
   END_VAR
   VAR_TEMP
      ErrorAbort : Bool;
   END_VAR
BEGIN

   IF (#Abort OR #Core.ReleasePending) AND #Core.Exec = 1 THEN
       #Core.Exec := 4;
       #Core.Step := 0;
       #Core.Dispatch := FALSE;
       #Core.EvAbort := TRUE;
   END_IF;
   #ErrorAbort := (#Abort OR #Core.ReleasePending) AND #Core.Exec = 3;
   #Core.EvAbortInError := #ErrorAbort AND NOT #Core.AbortPrev;
   #Core.AbortPrev := #ErrorAbort;
END_FUNCTION

FUNCTION "FRK_Route_CylinderCM" : Bool   // FC146, SCL
{ S7_Optimized_Access := 'TRUE' }
VERSION : 0.1
// stored: AutoNumber true, IsIECCheckEnabled false, SetENOAutomatically false, UDAEnableTagReadback false
   VAR_INPUT
      Request : "ST_HmiRequest";
   END_VAR
   VAR_IN_OUT
      Module : "FB_CylinderCM";
      Hal : "ST_CylinderHal";
      Report : "ST_ReleaseReport";
   END_VAR
   VAR_TEMP
      RouteMatched : Bool;
      Index : Int;
   END_VAR
BEGIN

   #FRK_Route_CylinderCM := FALSE;
   IF NOT "FRK_PathOwned"(OwnerPath := #Module.Status.Name, TargetPath := #Request.TargetPath) THEN
       RETURN;
   END_IF;
   IF #Request.TargetPath = STRING_TO_WSTRING(#Module.Status.Name) THEN
       FOR #Index := 1 TO 16 DO
           #Module.ManConditions[#Index].Used := FALSE;
       END_FOR;
       // ---- AUTHORED: OnManRelease
       "FRK_ManualCondition"(Conditions := #Module.ManConditions,
                             Slot := 1,
                             Value := 1,
                             Ok := #Hal.ExtendPermit,
                             Diag := #Hal.PermitDiagnostic,
                             Bypassable := FALSE);
       "FRK_ManualCondition"(Conditions := #Module.ManConditions,
                             Slot := 2,
                             Value := 2,
                             Ok := #Hal.RetractPermit,
                             Diag := #Hal.RetractDiagnostic,
                             Bypassable := FALSE);

       // ---- GENERATED: manual release end
       "FRK_ManualApply"(Core := #Module.Core,
                         Status := #Module.Status,
                         Request := #Request,
                         Commands := #Module.Catalog,
                         Count := #Module.CatalogCount,
                         Conditions := #Module.ManConditions,
                         Report := #Report,
                         Execute := #Module.Execute,
                         Command := #Module.Command,
                         ManualOwned := #Module.ManualOwned);
       #FRK_Route_CylinderCM := TRUE;
       RETURN;
   END_IF;
END_FUNCTION

FUNCTION "FRK_Route_PressDemoUnit" : Bool   // FC172, SCL
{ S7_Optimized_Access := 'TRUE' }
VERSION : 0.1
// stored: AutoNumber true, IsIECCheckEnabled false, SetENOAutomatically false, UDAEnableTagReadback false
   VAR_INPUT
      Request : "ST_HmiRequest";
   END_VAR
   VAR_IN_OUT
      Module : "FB_PressDemoUnit";
      Hal : "ST_PressDemoUnitHal";
      Report : "ST_ReleaseReport";
   END_VAR
   VAR_TEMP
      RouteMatched : Bool;
      Index : Int;
   END_VAR
BEGIN

   #FRK_Route_PressDemoUnit := FALSE;
   IF NOT "FRK_PathOwned"(OwnerPath := #Module.Status.Name, TargetPath := #Request.TargetPath) THEN
       RETURN;
   END_IF;
   "FRK_Release_PressDemoUnit"(Unit := #Module.Unit,
                               Hal := #Hal);
   "FRK_ManualCommon"(Core := #Module.Core,
                      Unit := #Module.Unit,
                      Status := #Module.Status,
                      Report := #Report);
   IF #Request.TargetPath = STRING_TO_WSTRING(#Module.Status.Name) THEN
       "FRK_ReleaseReason"(Report := #Report,
                           Description := WSTRING#'std.error.unsupportedHmiRequest',
                           Reason := 2008,
                           Path := STRING_TO_WSTRING(#Module.Status.Name),
                           Kind := 4);
       #FRK_Route_PressDemoUnit := TRUE;
       RETURN;
   END_IF;
   #RouteMatched := "FRK_Route_CylinderCM"(Module := #Module.PressRam, Hal := #Hal.PressRam, Request := #Request, Report := #Report);
   #FRK_Route_PressDemoUnit := #FRK_Route_PressDemoUnit OR #RouteMatched;
   #RouteMatched := "FRK_Route_CylinderCM"(Module := #Module.Door, Hal := #Hal.Door, Request := #Request, Report := #Report);
   #FRK_Route_PressDemoUnit := #FRK_Route_PressDemoUnit OR #RouteMatched;
   #RouteMatched := "FRK_Route_CylinderCM"(Module := #Module.PartSlide, Hal := #Hal.PartSlide, Request := #Request, Report := #Report);
   #FRK_Route_PressDemoUnit := #FRK_Route_PressDemoUnit OR #RouteMatched;
END_FUNCTION

FUNCTION "FRK_SeqAdvance" : Void   // FC132, SCL
{ S7_Optimized_Access := 'TRUE' }
VERSION : 0.1
// stored: AutoNumber true, IsIECCheckEnabled false, SetENOAutomatically false, UDAEnableTagReadback false
   VAR_INPUT
      Ok : Bool;
      OnAdvance : DInt;
   END_VAR
   VAR_IN_OUT
      Seq : "FRK_SequenceCtx";
   END_VAR
BEGIN

   "FRK_SeqSelect"(Seq := #Seq, AdvanceOk := #Ok, Jump1Ok := FALSE);
   "FRK_SeqRoute"(Seq := #Seq, OnAdvance := #OnAdvance, OnJump1 := -1);
END_FUNCTION

FUNCTION "FRK_SeqCommand" : Bool   // FC134, SCL
{ S7_Optimized_Access := 'TRUE' }
VERSION : 0.1
// stored: AutoNumber true, IsIECCheckEnabled false, SetENOAutomatically false, UDAEnableTagReadback false
   VAR_INPUT
      Value : DInt;
      Label : String;
      Ready : Bool;
      Done : Bool;
      Error : Bool;
      OwnFailure : Bool;
      Diagnostic : "ST_Diagnostic";
   END_VAR
   VAR_IN_OUT
      Seq : "FRK_SequenceCtx";
      Lease : "ST_SequenceCommandLease";
      Execute : Bool;
      Command : DInt;
   END_VAR
   VAR_TEMP
      WaitOk : Bool;
   END_VAR
BEGIN

   #FRK_SeqCommand := FALSE;
   IF NOT #Seq.Running OR #Seq.Error OR #Seq.OwnerIndex <= 0 OR #Seq.ChainIndex <= 0 THEN
       RETURN;
   END_IF;
   IF #Lease.Raised THEN
       IF #Lease.OwnerIndex <> #Seq.OwnerIndex OR #Lease.ChainIndex <> #Seq.ChainIndex OR #Lease.BranchIndex <> #Seq.BranchIndex
           OR #Lease.Step <> #Seq.Step OR #Command <> #Value THEN
           // Another chain owns this command; never borrow its Done result.
           #WaitOk := "FRK_SeqAwait"(Seq := #Seq, Label := 'std.release.commandOwned', Ok := FALSE);
           RETURN;
       END_IF;
       IF #Done THEN
           #FRK_SeqCommand := TRUE;
       ELSIF #Error THEN
           IF #OwnFailure THEN
               #Seq.CommandFailed := TRUE;
               #Seq.HandledDiagnostic := #Diagnostic;
           ELSE
               #Seq.Error := TRUE;
               #Seq.ErrorDiagnostic := #Diagnostic;
           END_IF;
           #Execute := FALSE;
       ELSE
           #WaitOk := "FRK_SeqAwait"(Seq := #Seq, Label := #Label, Ok := FALSE);
       END_IF;
   ELSIF #Ready AND #Lease.ReleasedScan <> #Seq.Scan THEN
       #Lease.OwnerIndex := #Seq.OwnerIndex;
       #Lease.ChainIndex := #Seq.ChainIndex;
       #Lease.BranchIndex := #Seq.BranchIndex;
       #Lease.Step := #Seq.Step;
       #Lease.Raised := TRUE;
       #Seq.CommandIssued := TRUE;
       #Command := #Value;
       #Execute := TRUE;
       #WaitOk := "FRK_SeqAwait"(Seq := #Seq, Label := #Label, Ok := FALSE);
   ELSE
       #WaitOk := "FRK_SeqAwait"(Seq := #Seq, Label := #Label, Ok := FALSE);
   END_IF;
END_FUNCTION

FUNCTION "FRK_SeqCycleEnd" : Void   // FC126, SCL
{ S7_Optimized_Access := 'TRUE' }
VERSION : 0.1
// stored: AutoNumber true, IsIECCheckEnabled false, SetENOAutomatically false, UDAEnableTagReadback false
   VAR_IN_OUT
      Seq : "FRK_SequenceCtx";
   END_VAR
BEGIN

   #Seq.StartLatched := FALSE;
END_FUNCTION

FUNCTION "FRK_SeqHandled" : Void   // FC140, SCL
{ S7_Optimized_Access := 'TRUE' }
VERSION : 0.1
// stored: AutoNumber true, IsIECCheckEnabled false, SetENOAutomatically false, UDAEnableTagReadback false
   VAR_IN_OUT
      Seq : "FRK_SequenceCtx";
      ChildCore : "FRK_Core";
   END_VAR
BEGIN

   // The owning step reports this occurrence through the closed AUTO_RESET
   // path. Ordinary child faults retain their MANUAL_RESET capture.
   IF #Seq.CommandFailed THEN
       #ChildCore.FaultHandled := TRUE;
   END_IF;
END_FUNCTION

FUNCTION "FRK_SeqLease" : Void   // FC133, SCL
{ S7_Optimized_Access := 'TRUE' }
VERSION : 0.1
// stored: AutoNumber true, IsIECCheckEnabled false, SetENOAutomatically false, UDAEnableTagReadback false
   VAR_IN_OUT
      Seq : "FRK_SequenceCtx";
      Lease : "ST_SequenceCommandLease";
      Execute : Bool;
   END_VAR
BEGIN

   IF #Lease.Raised AND #Lease.OwnerIndex > 0 AND #Lease.ChainIndex > 0
       AND #Lease.OwnerIndex = #Seq.OwnerIndex AND #Lease.ChainIndex = #Seq.ChainIndex
       AND #Lease.BranchIndex = #Seq.BranchIndex THEN
       IF NOT #Seq.Running OR #Seq.Error OR #Seq.Restart OR #Lease.Step <> #Seq.Step THEN
           #Execute := FALSE;
           #Lease.Raised := FALSE;
           #Lease.ReleasedScan := #Seq.Scan;
       END_IF;
   END_IF;
END_FUNCTION

FUNCTION "FRK_SeqMessage" : Void   // FC144, SCL
{ S7_Optimized_Access := 'TRUE' }
VERSION : 0.1
// stored: AutoNumber true, IsIECCheckEnabled false, SetENOAutomatically false, UDAEnableTagReadback false
   VAR_INPUT
      Diag : "ST_Diagnostic";
   END_VAR
   VAR_IN_OUT
      Seq : "FRK_SequenceCtx";
      AlarmLog : "FRK_AlarmLog";
   END_VAR
   VAR_TEMP
      Slot : Int;
      Gone : Bool;
   END_VAR
BEGIN

   IF #Seq.Warned THEN
       RETURN;
   END_IF;
   #Slot := "FRK_AlarmRaise"(AlarmLog := #AlarmLog, Diag := #Diag, ResetClass := 0);
   IF #Slot > 0 THEN
       #Gone := "FRK_AlarmGone"(AlarmLog := #AlarmLog, Slot := #Slot);
       #Seq.Warned := TRUE;
   END_IF;
END_FUNCTION

FUNCTION "FRK_SeqOnce" : Bool   // FC143, SCL
{ S7_Optimized_Access := 'TRUE' }
VERSION : 0.1
// stored: AutoNumber true, IsIECCheckEnabled false, SetENOAutomatically false, UDAEnableTagReadback false
   VAR_INPUT
      Enable : Bool;
      Token : DInt;
   END_VAR
   VAR_IN_OUT
      Seq : "FRK_SequenceCtx";
   END_VAR
BEGIN

   #FRK_SeqOnce := #Enable AND #Seq.Running AND NOT #Seq.Error
   AND (#Seq.EventVisit <> #Seq.Visit OR #Seq.EventToken <> #Token);
   IF #FRK_SeqOnce THEN
       #Seq.EventVisit := #Seq.Visit;
       #Seq.EventToken := #Token;
   END_IF;
END_FUNCTION

FUNCTION "FRK_SeqSelect" : Void   // FC139, SCL
{ S7_Optimized_Access := 'TRUE' }
VERSION : 0.1
// stored: AutoNumber true, IsIECCheckEnabled false, SetENOAutomatically false, UDAEnableTagReadback false
   VAR_INPUT
      AdvanceOk : Bool;
      Jump1Ok : Bool;
   END_VAR
   VAR_IN_OUT
      Seq : "FRK_SequenceCtx";
   END_VAR
BEGIN

   #Seq.RetVal := 0;
   IF NOT #Seq.Running OR #Seq.Error THEN
       RETURN;
   END_IF;
   IF #AdvanceOk THEN
       #Seq.RetVal := 1;
   ELSIF #Jump1Ok THEN
       #Seq.RetVal := 2;
   END_IF;
END_FUNCTION

FUNCTION "FRK_SetBoot" : Void   // FC117, SCL
{ S7_Optimized_Access := 'TRUE' }
VERSION : 0.1
// stored: AutoNumber true, IsIECCheckEnabled false, SetENOAutomatically false, UDAEnableTagReadback false
   VAR_INPUT
      Startup : Bool;
   END_VAR
   VAR_TEMP
      RootIndex : Int;
      Slot : Int;
   END_VAR
BEGIN

   IF NOT #Startup THEN
       RETURN;
   END_IF;
   IF "FRK_SetStore".SchemaVersion <> 1 THEN
       FOR #RootIndex := 1 TO 1 DO
           IF "FRK_SetStore".SchemaVersion <> 0 THEN
               "FRK_ConfigLoss"(RootIndex := #RootIndex,
                                Scope := "FRK_SetStore".Sets[#RootIndex, 1].Info.RootIdentity);
           END_IF;
           FOR #Slot := 1 TO 4 DO
               "FRK_SetStore".Sets[#RootIndex, #Slot].Info.Used := FALSE;
           END_FOR;
       END_FOR;
       "FRK_SetStore".SchemaVersion := 1;
   END_IF;
END_FUNCTION

FUNCTION "FRK_SetCheck" : Int   // FC107, SCL
{ S7_Optimized_Access := 'TRUE' }
VERSION : 0.1
// stored: AutoNumber true, IsIECCheckEnabled false, SetENOAutomatically false, UDAEnableTagReadback false
   VAR_INPUT
      RootIndex : Int;
      Scope : String;
      Access : "FRK_Access";
      Ready : Bool;
      WriteAccess : Bool;
   END_VAR
   VAR_TEMP
      Index : Int;
      Ok : Bool;
   END_VAR
BEGIN

   #FRK_SetCheck := 0;
   "FRK_SetRuntime".Work[#RootIndex].RejectScope := #Scope;
   "FRK_SetRuntime".Work[#RootIndex].RejectKey := "FRK_ConfigScratch".Entry.WriteKey;
   #Index := "FRK_SetRecord"(RootIndex := #RootIndex, Scope := #Scope, WriteKey := "FRK_ConfigScratch".Entry.WriteKey);
   IF #Index = 0 THEN
       RETURN;
   END_IF;
   IF #Access.CurrentLevel < MAX(IN1 := #Access.Policy.Required[0], IN2 := "FRK_ConfigScratch".MinRead) THEN
       RETURN;
   END_IF;
   IF #WriteAccess THEN
       IF #Access.CurrentLevel < MAX(IN1 := #Access.Policy.Required[1], IN2 := "FRK_ConfigScratch".MinWrite) THEN
           RETURN;
       END_IF;
       IF "FRK_ConfigScratch".Entry.RequiresReady AND NOT #Ready THEN
           RETURN;
       END_IF;
   END_IF;
   IF "FRK_SetRuntime".Work[#RootIndex].Payload.Records[#Index].Revision <> "FRK_ConfigScratch".Entry.WriteRevision
       OR "FRK_SetRuntime".Work[#RootIndex].Payload.Records[#Index].Kind <> "FRK_ConfigScratch".Entry.ConfigKind
       OR "FRK_SetRuntime".Work[#RootIndex].Payload.Records[#Index].ValueType <> "FRK_ConfigScratch".Entry.ValueType THEN
       RETURN;
   END_IF;
   #Ok := "FRK_ConfigDecode"(Text := STRING_TO_WSTRING("FRK_SetRuntime".Work[#RootIndex].Payload.Records[#Index].ValueText), Storage := "FRK_ConfigScratch".Storage,
                             Minimum := "FRK_ConfigScratch".Minimum, Maximum := "FRK_ConfigScratch".Maximum, MaxLength := "FRK_ConfigScratch".MaxLength, Value := "FRK_ConfigScratch".Value);
   IF NOT #Ok THEN
       RETURN;
   END_IF;
   // Existing keyed slots are reserved before commit: commit cannot allocate.
   IF #WriteAccess AND "FRK_ConfigFind"(Scope := #Scope, Key := "FRK_ConfigScratch".Entry.WriteKey, ModelCode := "FRK_SetRuntime".Work[#RootIndex].Payload.Info.ModelCode) = 0 THEN
       RETURN;
   END_IF;
   "FRK_SetRuntime".Work[#RootIndex].Seen[#Index] := TRUE;
   "FRK_SetRuntime".Work[#RootIndex].Matched := "FRK_SetRuntime".Work[#RootIndex].Matched + 1;
   #FRK_SetCheck := #Index;
END_FUNCTION

FUNCTION "FRK_SetFind" : Int   // FC104, SCL
{ S7_Optimized_Access := 'TRUE' }
VERSION : 0.1
// Deployment-sized keyed set storage; validation belongs to the typed walk.
// stored: AutoNumber true, IsIECCheckEnabled false, SetENOAutomatically false, UDAEnableTagReadback false
   VAR_INPUT
      RootIndex : Int;
      SetName : String;
   END_VAR
   VAR_TEMP
      Index : Int;
   END_VAR
BEGIN

   #FRK_SetFind := 0;
   FOR #Index := 1 TO 4 DO
       IF "FRK_SetStore".Sets[#RootIndex, #Index].Info.Used AND "FRK_SetStore".Sets[#RootIndex, #Index].Info.SetName = #SetName THEN
           #FRK_SetFind := #Index;
           RETURN;
       END_IF;
   END_FOR;
END_FUNCTION

FUNCTION "FRK_SetIdentity" : Void   // FC1, SCL
{ S7_Optimized_Access := 'TRUE' }
VERSION : 0.1
// Generated registry services v0.1; compact rows contain no operator strings.
// stored: AutoNumber true, IsIECCheckEnabled false, SetENOAutomatically false, UDAEnableTagReadback false
   VAR_INPUT
      InstancePath : WString;
      ModuleType : DInt;
      TypeId : DInt;
      Capabilities : DWord;
      ParentIndex : DInt;
      TypeKey : String;
   END_VAR
   VAR_IN_OUT
      Core : "FRK_Core";
      Status : "ST_ModuleStatus";
   END_VAR
   VAR_TEMP
      Identity : String[254];
      QuotePos : Int;
      RowIndex : DInt;
   END_VAR
BEGIN

   #Core.Named := TRUE;
   #Core.RegIndex := 0;
   IF "FRK_Registry".Fault OR "FRK_Registry".Count < 0 OR "FRK_Registry".Count > 4
       OR #ParentIndex < 0 OR #ParentIndex > "FRK_Registry".Count OR #ParentIndex > 4 THEN
       "FRK_Registry".Fault := TRUE;
       RETURN;
   END_IF;
   IF #ParentIndex > 0 THEN
       IF NOT "FRK_Registry".Rows[#ParentIndex].Valid THEN
           "FRK_Registry".Fault := TRUE;
           RETURN;
       END_IF;
   END_IF;
   IF LEN(#InstancePath) > 254 THEN
       "FRK_Registry".Fault := TRUE;
       RETURN;
   END_IF;
   #Identity := WSTRING_TO_STRING(#InstancePath);
   #QuotePos := FIND(IN1 := #Identity, IN2 := '"');
   WHILE #QuotePos > 0 DO
       #Identity := DELETE(IN := #Identity, L := 1, P := #QuotePos);
       #QuotePos := FIND(IN1 := #Identity, IN2 := '"');
   END_WHILE;
   IF LEN(#Identity) > 80 OR LEN(#Identity) = 0 OR "FRK_Registry".Count >= 4 THEN
       "FRK_Registry".Fault := TRUE;
       RETURN;
   END_IF;
   "FRK_Registry".Count := "FRK_Registry".Count + 1;
   #RowIndex := "FRK_Registry".Count;
   #Core.RegIndex := #RowIndex;
   #Core.ParentIndex := #ParentIndex;
   #Core.ModuleType := #ModuleType;
   #Status.Name := #Identity;
   #Status.TypeKey := #TypeKey;
   #Status.ModuleType := #ModuleType;
   #Status.TileEnable := TRUE;
   "FRK_Registry".Rows[#RowIndex].Valid := TRUE;
   "FRK_Registry".Rows[#RowIndex].Parent := #ParentIndex;
   "FRK_Registry".Rows[#RowIndex].ModuleType := #ModuleType;
   "FRK_Registry".Rows[#RowIndex].TypeId := #TypeId;
   "FRK_Registry".Rows[#RowIndex].Capabilities := #Capabilities;
END_FUNCTION

FUNCTION "FRK_SetImport" : Bool   // FC112, SCL
{ S7_Optimized_Access := 'TRUE' }
VERSION : 0.1
// stored: AutoNumber true, IsIECCheckEnabled false, SetENOAutomatically false, UDAEnableTagReadback false
   VAR_INPUT
      RootIndex : Int;
      Request : "ST_HmiRequest";
   END_VAR
   VAR_TEMP
      Ok : Bool;
      Index : Int;
   END_VAR
BEGIN

   #FRK_SetImport := FALSE;
   IF #Request.IntValue <> 0 AND #Request.IntValue <> 1 THEN
       RETURN;
   END_IF;
   IF #Request.NameValue <> '' OR #Request.TargetPath <> WSTRING#'' OR #Request.DurationMs <> 0 THEN
       RETURN;
   END_IF;
   #Ok := "FRK_JsonPut"(Text := #Request.TextValue, Line := "FRK_SetRuntime".Work[#RootIndex].Piece);
   IF NOT #Ok THEN
       RETURN;
   END_IF;
   IF #Request.IntValue = 1 THEN
       #FRK_SetImport := NOT #Request.BoolValue;
       RETURN;
   END_IF;
   "FRK_SetRuntime".Work[#RootIndex].Line := "FRK_SetRuntime".Work[#RootIndex].Piece;
   "FRK_SetRuntime".Work[#RootIndex].Piece := WSTRING#'';
   #Ok := "FRK_JsonParse"(Line := "FRK_SetRuntime".Work[#RootIndex].Line, Fields := "FRK_SetRuntime".Work[#RootIndex].Fields, Count := "FRK_SetRuntime".Work[#RootIndex].FieldCount);
   IF NOT #Ok THEN
       RETURN;
   END_IF;
   IF NOT "FRK_SetRuntime".Work[#RootIndex].Importing THEN
       #Ok := "FRK_JsonReadHeader"(Count := "FRK_SetRuntime".Work[#RootIndex].FieldCount,
                                   Fields := "FRK_SetRuntime".Work[#RootIndex].Fields,
                                   Data := "FRK_SetRuntime".Work[#RootIndex].Payload.Info);
       IF NOT #Ok OR #Request.BoolValue THEN
           RETURN;
       END_IF;
       "FRK_SetRuntime".Work[#RootIndex].Payload.Info.Used := TRUE;
       "FRK_SetRuntime".Work[#RootIndex].Received := 0;
       "FRK_SetRuntime".Work[#RootIndex].Importing := TRUE;
   ELSE
       #Index := "FRK_SetRuntime".Work[#RootIndex].Received + 1;
       IF #Index > 3 OR #Index > "FRK_SetRuntime".Work[#RootIndex].Payload.Info.RecordCount THEN
           RETURN;
       END_IF;
       #Ok := "FRK_JsonReadRecord"(Count := "FRK_SetRuntime".Work[#RootIndex].FieldCount,
                                   Fields := "FRK_SetRuntime".Work[#RootIndex].Fields,
                                   Data := "FRK_SetRuntime".Work[#RootIndex].Payload.Records[#Index]);
       IF NOT #Ok THEN
           RETURN;
       END_IF;
       "FRK_SetRuntime".Work[#RootIndex].Received := #Index;
   END_IF;
   IF #Request.BoolValue THEN
       "FRK_SetRuntime".Work[#RootIndex].Importing := FALSE;
       IF "FRK_SetRuntime".Work[#RootIndex].Received <> "FRK_SetRuntime".Work[#RootIndex].Payload.Info.RecordCount THEN
           RETURN;
       END_IF;
   END_IF;
   #FRK_SetImport := TRUE;
END_FUNCTION

FUNCTION "FRK_SetRecord" : Int   // FC106, SCL
{ S7_Optimized_Access := 'TRUE' }
VERSION : 0.1
// stored: AutoNumber true, IsIECCheckEnabled false, SetENOAutomatically false, UDAEnableTagReadback false
   VAR_INPUT
      RootIndex : Int;
      Scope : String;
      WriteKey : String;
   END_VAR
   VAR_TEMP
      Index : Int;
   END_VAR
BEGIN

   #FRK_SetRecord := 0;
   FOR #Index := 1 TO "FRK_SetRuntime".Work[#RootIndex].Payload.Info.RecordCount DO
       IF "FRK_SetRuntime".Work[#RootIndex].Payload.Records[#Index].Scope = #Scope AND "FRK_SetRuntime".Work[#RootIndex].Payload.Records[#Index].WriteKey = #WriteKey THEN
           #FRK_SetRecord := #Index;
           RETURN;
       END_IF;
   END_FOR;
END_FUNCTION

FUNCTION "FRK_SetResult" : Void   // FC116, SCL
{ S7_Optimized_Access := 'TRUE' }
VERSION : 0.1
// stored: AutoNumber true, IsIECCheckEnabled false, SetENOAutomatically false, UDAEnableTagReadback false
   VAR_INPUT
      Request : "ST_HmiRequest";
      Response : "ST_HmiResponse";
      Scope : String;
      RootIndex : Int;
   END_VAR
   VAR_IN_OUT
      Persist : "ST_ConfigPersistStatus";
      AlarmLog : "FRK_AlarmLog";
   END_VAR
   VAR_TEMP
      Diag : "ST_Diagnostic";
      Slot : Int;
      Ok : Bool;
   END_VAR
BEGIN

   IF #Request.Kind <> 29 THEN
       RETURN;
   END_IF;
   IF NOT #Response.Accepted THEN
       #Persist.LastRejectScope := "FRK_SetRuntime".Work[#RootIndex].RejectScope;
       #Persist.LastRejectKey := "FRK_SetRuntime".Work[#RootIndex].RejectKey;
   END_IF;
   #Diag := "FRK_UnitScratch".EmptyDiagnostic;
   #Diag.SourcePath := STRING_TO_WSTRING(#Scope);
   IF #Response.Accepted THEN
       #Diag.ReasonCode := 2043;
       #Diag.Description := WSTRING#'std.event.configSetApplied';
   ELSE
       #Diag.ReasonCode := 2042;
       #Diag.Description := WSTRING#'std.error.configSetRejected';
       #Diag.SourcePath := STRING_TO_WSTRING(#Persist.LastRejectScope);
   END_IF;
   #Slot := "FRK_AlarmRaise"(AlarmLog := #AlarmLog, Diag := #Diag, ResetClass := 0);
   IF #Slot > 0 THEN
       #Ok := "FRK_AlarmGone"(AlarmLog := #AlarmLog, Slot := #Slot);
   END_IF;
END_FUNCTION

FUNCTION "FRK_SetShape" : Bool   // FC111, SCL
{ S7_Optimized_Access := 'TRUE' }
VERSION : 0.1
// stored: AutoNumber true, IsIECCheckEnabled false, SetENOAutomatically false, UDAEnableTagReadback false
   VAR_INPUT
      RootIndex : Int;
      RootIdentity : String;
   END_VAR
   VAR_TEMP
      Index : Int;
      Other : Int;
      ModelIndex : Int;
      KnownModel : Bool;
   END_VAR
BEGIN

   #FRK_SetShape := FALSE;
   IF NOT "FRK_SetRuntime".Work[#RootIndex].Payload.Info.Used OR "FRK_SetRuntime".Work[#RootIndex].Payload.Info.RootIdentity <> #RootIdentity
       OR "FRK_SetRuntime".Work[#RootIndex].Payload.Info.SetSchema <> 1 OR "FRK_SetRuntime".Work[#RootIndex].Payload.Info.ConfigRev = 0
       OR LEN("FRK_SetRuntime".Work[#RootIndex].Payload.Info.SetName) = 0
       OR "FRK_SetRuntime".Work[#RootIndex].Payload.Info.RecordCount < 1 OR "FRK_SetRuntime".Work[#RootIndex].Payload.Info.RecordCount > 3 THEN
       RETURN;
   END_IF;
   IF "FRK_SetRuntime".Work[#RootIndex].Payload.Info.Kind = 0 THEN
       #KnownModel := FALSE;
       IF NOT #KnownModel THEN
           RETURN;
       END_IF;
   ELSIF "FRK_SetRuntime".Work[#RootIndex].Payload.Info.Kind <> 1 OR "FRK_SetRuntime".Work[#RootIndex].Payload.Info.ModelCode <> '' THEN
       RETURN;
   END_IF;
   FOR #Index := 1 TO "FRK_SetRuntime".Work[#RootIndex].Payload.Info.RecordCount DO
       "FRK_SetRuntime".Work[#RootIndex].RejectScope := "FRK_SetRuntime".Work[#RootIndex].Payload.Records[#Index].Scope;
       "FRK_SetRuntime".Work[#RootIndex].RejectKey := "FRK_SetRuntime".Work[#RootIndex].Payload.Records[#Index].WriteKey;
       IF "FRK_SetRuntime".Work[#RootIndex].Payload.Records[#Index].Kind <> "FRK_SetRuntime".Work[#RootIndex].Payload.Info.Kind THEN
           RETURN;
       END_IF;
       FOR #Other := 1 TO #Index - 1 DO
           IF "FRK_SetRuntime".Work[#RootIndex].Payload.Records[#Other].Scope = "FRK_SetRuntime".Work[#RootIndex].Payload.Records[#Index].Scope
               AND "FRK_SetRuntime".Work[#RootIndex].Payload.Records[#Other].WriteKey = "FRK_SetRuntime".Work[#RootIndex].Payload.Records[#Index].WriteKey THEN
               RETURN;
           END_IF;
       END_FOR;
   END_FOR;
   #FRK_SetShape := TRUE;
END_FUNCTION

FUNCTION "FRK_SetSlot" : Int   // FC105, SCL
{ S7_Optimized_Access := 'TRUE' }
VERSION : 0.1
// stored: AutoNumber true, IsIECCheckEnabled false, SetENOAutomatically false, UDAEnableTagReadback false
   VAR_INPUT
      RootIndex : Int;
      SetName : String;
   END_VAR
   VAR_TEMP
      Index : Int;
   END_VAR
BEGIN

   #FRK_SetSlot := "FRK_SetFind"(RootIndex := #RootIndex, SetName := #SetName);
   IF #FRK_SetSlot <> 0 THEN
       RETURN;
   END_IF;
   FOR #Index := 1 TO 4 DO
       IF NOT "FRK_SetStore".Sets[#RootIndex, #Index].Info.Used THEN
           #FRK_SetSlot := #Index;
           RETURN;
       END_IF;
   END_FOR;
END_FUNCTION

FUNCTION "FRK_SetValidateBegin" : Void   // FC114, SCL
{ S7_Optimized_Access := 'TRUE' }
VERSION : 0.1
// stored: AutoNumber true, IsIECCheckEnabled false, SetENOAutomatically false, UDAEnableTagReadback false
   VAR_INPUT
      RootIndex : Int;
   END_VAR
   VAR_TEMP
      Index : Int;
   END_VAR
BEGIN

   "FRK_SetRuntime".Work[#RootIndex].Matched := 0;
   FOR #Index := 1 TO 3 DO
       "FRK_SetRuntime".Work[#RootIndex].Seen[#Index] := FALSE;
   END_FOR;
END_FUNCTION

FUNCTION "FRK_SetValidateEnd" : Bool   // FC115, SCL
{ S7_Optimized_Access := 'TRUE' }
VERSION : 0.1
// stored: AutoNumber true, IsIECCheckEnabled false, SetENOAutomatically false, UDAEnableTagReadback false
   VAR_INPUT
      RootIndex : Int;
   END_VAR
   VAR_TEMP
      Index : Int;
   END_VAR
BEGIN

   #FRK_SetValidateEnd := FALSE;
   FOR #Index := 1 TO "FRK_SetRuntime".Work[#RootIndex].Payload.Info.RecordCount DO
       IF NOT "FRK_SetRuntime".Work[#RootIndex].Seen[#Index] THEN
           "FRK_SetRuntime".Work[#RootIndex].RejectScope := "FRK_SetRuntime".Work[#RootIndex].Payload.Records[#Index].Scope;
           "FRK_SetRuntime".Work[#RootIndex].RejectKey := "FRK_SetRuntime".Work[#RootIndex].Payload.Records[#Index].WriteKey;
           RETURN;
       END_IF;
   END_FOR;
   #FRK_SetValidateEnd := "FRK_SetRuntime".Work[#RootIndex].Matched = "FRK_SetRuntime".Work[#RootIndex].Payload.Info.RecordCount;
END_FUNCTION

FUNCTION "FRK_Sha256Pin" : Bool   // FC39, SCL
{ S7_Optimized_Access := 'TRUE' }
VERSION : 0.1
// Core section 7.7 prototype: private retained provider injection and independent root sessions.
//  User records are salted Core-compatible hashes, never commissioning plaintext.
// stored: AutoNumber true, IsIECCheckEnabled false, SetENOAutomatically false, UDAEnableTagReadback false
   VAR_INPUT
      Size : DInt;
   END_VAR
   VAR_IN_OUT
      Data : Array[0..47] of Byte;
      Digest : Array[0..31] of Byte;
   END_VAR
   VAR_TEMP
      BlockBytes : Array[0..63] of Byte;
      Words : Array[0..63] of DWord;
      Hash : Array[0..7] of DWord;
      Index : DInt;
      "A" : DWord;
      "B" : DWord;
      C : DWord;
      D : DWord;
      "E" : DWord;
      F : DWord;
      G : DWord;
      H : DWord;
      S0 : DWord;
      S1 : DWord;
      T1 : DWord;
      T2 : DWord;
      K : Array[0..63] of DWord;
   END_VAR
BEGIN

   #FRK_Sha256Pin := FALSE;
   #K[0] := DWORD#16#428A2F98;
   #K[1] := DWORD#16#71374491;
   #K[2] := DWORD#16#B5C0FBCF;
   #K[3] := DWORD#16#E9B5DBA5;
   #K[4] := DWORD#16#3956C25B;
   #K[5] := DWORD#16#59F111F1;
   #K[6] := DWORD#16#923F82A4;
   #K[7] := DWORD#16#AB1C5ED5;
   #K[8] := DWORD#16#D807AA98;
   #K[9] := DWORD#16#12835B01;
   #K[10] := DWORD#16#243185BE;
   #K[11] := DWORD#16#550C7DC3;
   #K[12] := DWORD#16#72BE5D74;
   #K[13] := DWORD#16#80DEB1FE;
   #K[14] := DWORD#16#9BDC06A7;
   #K[15] := DWORD#16#C19BF174;
   #K[16] := DWORD#16#E49B69C1;
   #K[17] := DWORD#16#EFBE4786;
   #K[18] := DWORD#16#0FC19DC6;
   #K[19] := DWORD#16#240CA1CC;
   #K[20] := DWORD#16#2DE92C6F;
   #K[21] := DWORD#16#4A7484AA;
   #K[22] := DWORD#16#5CB0A9DC;
   #K[23] := DWORD#16#76F988DA;
   #K[24] := DWORD#16#983E5152;
   #K[25] := DWORD#16#A831C66D;
   #K[26] := DWORD#16#B00327C8;
   #K[27] := DWORD#16#BF597FC7;
   #K[28] := DWORD#16#C6E00BF3;
   #K[29] := DWORD#16#D5A79147;
   #K[30] := DWORD#16#06CA6351;
   #K[31] := DWORD#16#14292967;
   #K[32] := DWORD#16#27B70A85;
   #K[33] := DWORD#16#2E1B2138;
   #K[34] := DWORD#16#4D2C6DFC;
   #K[35] := DWORD#16#53380D13;
   #K[36] := DWORD#16#650A7354;
   #K[37] := DWORD#16#766A0ABB;
   #K[38] := DWORD#16#81C2C92E;
   #K[39] := DWORD#16#92722C85;
   #K[40] := DWORD#16#A2BFE8A1;
   #K[41] := DWORD#16#A81A664B;
   #K[42] := DWORD#16#C24B8B70;
   #K[43] := DWORD#16#C76C51A3;
   #K[44] := DWORD#16#D192E819;
   #K[45] := DWORD#16#D6990624;
   #K[46] := DWORD#16#F40E3585;
   #K[47] := DWORD#16#106AA070;
   #K[48] := DWORD#16#19A4C116;
   #K[49] := DWORD#16#1E376C08;
   #K[50] := DWORD#16#2748774C;
   #K[51] := DWORD#16#34B0BCB5;
   #K[52] := DWORD#16#391C0CB3;
   #K[53] := DWORD#16#4ED8AA4A;
   #K[54] := DWORD#16#5B9CCA4F;
   #K[55] := DWORD#16#682E6FF3;
   #K[56] := DWORD#16#748F82EE;
   #K[57] := DWORD#16#78A5636F;
   #K[58] := DWORD#16#84C87814;
   #K[59] := DWORD#16#8CC70208;
   #K[60] := DWORD#16#90BEFFFA;
   #K[61] := DWORD#16#A4506CEB;
   #K[62] := DWORD#16#BEF9A3F7;
   #K[63] := DWORD#16#C67178F2;
   FOR #Index := 0 TO 31 DO
       #Digest[#Index] := 0;
   END_FOR;
   IF #Size < 0 OR #Size > 48 THEN
       RETURN;
   END_IF;
   // Authentication messages fit exactly one SHA-256 block.
   FOR #Index := 0 TO 63 DO
       #BlockBytes[#Index] := 0;
   END_FOR;
   FOR #Index := 0 TO #Size - 1 DO
       #BlockBytes[#Index] := #Data[#Index];
   END_FOR;
   #BlockBytes[#Size] := BYTE#16#80;
   #BlockBytes[62] := DWORD_TO_BYTE(SHR(IN := DINT_TO_DWORD(#Size * 8), N := 8));
   #BlockBytes[63] := DINT_TO_BYTE(#Size * 8);
   #Hash[0] := DWORD#16#6A09E667;
   #Hash[1] := DWORD#16#BB67AE85;
   #Hash[2] := DWORD#16#3C6EF372;
   #Hash[3] := DWORD#16#A54FF53A;
   #Hash[4] := DWORD#16#510E527F;
   #Hash[5] := DWORD#16#9B05688C;
   #Hash[6] := DWORD#16#1F83D9AB;
   #Hash[7] := DWORD#16#5BE0CD19;
   FOR #Index := 0 TO 15 DO
       #Words[#Index] := SHL(IN := BYTE_TO_DWORD(#BlockBytes[4 * #Index]), N := 24)
       OR SHL(IN := BYTE_TO_DWORD(#BlockBytes[4 * #Index + 1]), N := 16)
       OR SHL(IN := BYTE_TO_DWORD(#BlockBytes[4 * #Index + 2]), N := 8)
       OR BYTE_TO_DWORD(#BlockBytes[4 * #Index + 3]);
   END_FOR;
   FOR #Index := 16 TO 63 DO
       #S0 := ROR(IN := #Words[#Index - 15], N := 7) XOR ROR(IN := #Words[#Index - 15], N := 18) XOR SHR(IN := #Words[#Index - 15], N := 3);
       #S1 := ROR(IN := #Words[#Index - 2], N := 17) XOR ROR(IN := #Words[#Index - 2], N := 19) XOR SHR(IN := #Words[#Index - 2], N := 10);
       #Words[#Index] := UDINT_TO_DWORD(ULINT_TO_UDINT(UDINT_TO_ULINT(DWORD_TO_UDINT(#Words[#Index - 16])) + UDINT_TO_ULINT(DWORD_TO_UDINT(#S0)) + UDINT_TO_ULINT(DWORD_TO_UDINT(#Words[#Index - 7])) + UDINT_TO_ULINT(DWORD_TO_UDINT(#S1))));
   END_FOR;
   #A := #Hash[0];
   #B := #Hash[1];
   #C := #Hash[2];
   #D := #Hash[3];
   #E := #Hash[4];
   #F := #Hash[5];
   #G := #Hash[6];
   #H := #Hash[7];
   FOR #Index := 0 TO 63 DO
       #S1 := ROR(IN := #E, N := 6) XOR ROR(IN := #E, N := 11) XOR ROR(IN := #E, N := 25);
       #T1 := UDINT_TO_DWORD(ULINT_TO_UDINT(UDINT_TO_ULINT(DWORD_TO_UDINT(#H)) + UDINT_TO_ULINT(DWORD_TO_UDINT(#S1)) + UDINT_TO_ULINT(DWORD_TO_UDINT((#E AND #F) XOR ((NOT #E) AND #G))) + UDINT_TO_ULINT(DWORD_TO_UDINT(#K[#Index])) + UDINT_TO_ULINT(DWORD_TO_UDINT(#Words[#Index]))));
       #S0 := ROR(IN := #A, N := 2) XOR ROR(IN := #A, N := 13) XOR ROR(IN := #A, N := 22);
       #T2 := UDINT_TO_DWORD(ULINT_TO_UDINT(UDINT_TO_ULINT(DWORD_TO_UDINT(#S0)) + UDINT_TO_ULINT(DWORD_TO_UDINT((#A AND #B) XOR (#A AND #C) XOR (#B AND #C)))));
       #H := #G;
       #G := #F;
       #F := #E;
       #E := UDINT_TO_DWORD(ULINT_TO_UDINT(UDINT_TO_ULINT(DWORD_TO_UDINT(#D)) + UDINT_TO_ULINT(DWORD_TO_UDINT(#T1))));
       #D := #C;
       #C := #B;
       #B := #A;
       #A := UDINT_TO_DWORD(ULINT_TO_UDINT(UDINT_TO_ULINT(DWORD_TO_UDINT(#T1)) + UDINT_TO_ULINT(DWORD_TO_UDINT(#T2))));
   END_FOR;
   #Words[0] := #A;
   #Words[1] := #B;
   #Words[2] := #C;
   #Words[3] := #D;
   #Words[4] := #E;
   #Words[5] := #F;
   #Words[6] := #G;
   #Words[7] := #H;
   FOR #Index := 0 TO 7 DO
       #Hash[#Index] := UDINT_TO_DWORD(ULINT_TO_UDINT(UDINT_TO_ULINT(DWORD_TO_UDINT(#Hash[#Index])) + UDINT_TO_ULINT(DWORD_TO_UDINT(#Words[#Index]))));
       #Digest[4 * #Index] := DWORD_TO_BYTE(SHR(IN := #Hash[#Index], N := 24));
       #Digest[4 * #Index + 1] := DWORD_TO_BYTE(SHR(IN := #Hash[#Index], N := 16));
       #Digest[4 * #Index + 2] := DWORD_TO_BYTE(SHR(IN := #Hash[#Index], N := 8));
       #Digest[4 * #Index + 3] := DWORD_TO_BYTE(#Hash[#Index]);
   END_FOR;
   FOR #Index := 0 TO 63 DO
       #BlockBytes[#Index] := 0;
       #Words[#Index] := 0;
   END_FOR;
   #FRK_Sha256Pin := TRUE;
END_FUNCTION

FUNCTION "FRK_Start" : Void   // FC14, SCL
{ S7_Optimized_Access := 'TRUE' }
VERSION : 0.1
// stored: AutoNumber true, IsIECCheckEnabled false, SetENOAutomatically false, UDAEnableTagReadback false
   VAR_INPUT
      Supported : Bool;
      Timeout : Time;
      Label : String;
   END_VAR
   VAR_IN_OUT
      Core : "FRK_Core";
      Status : "ST_ModuleStatus";
   END_VAR
BEGIN

   #Core.CommandLabel := #Label;
   IF NOT #Supported THEN
       "FRK_Fault"(Core := #Core,
                   Status := #Status,
                   ReasonCode := 2008,
                   Description := WSTRING#'fraktal.command.unsupported');
   ELSIF #Timeout <= T#0ms THEN
       "FRK_Fault"(Core := #Core,
                   Status := #Status,
                   ReasonCode := 2004,
                   Description := WSTRING#'fraktal.command.timeout.invalid');
   ELSE
       #Core.TimeoutMs := DINT_TO_UDINT(TIME_TO_DINT(#Timeout));
   END_IF;
END_FUNCTION

FUNCTION "FRK_State" : Bool   // FC21, SCL
{ S7_Optimized_Access := 'TRUE' }
VERSION : 0.1
// stored: AutoNumber true, IsIECCheckEnabled false, SetENOAutomatically false, UDAEnableTagReadback false
   VAR_INPUT
      Idx : Int;
      Key : String;
      Ok : Bool;
   END_VAR
   VAR_IN_OUT
      Flags : Array[1..12] of "ST_StateFlag";
      Count : Int;
      Touched : Array[1..12] of Bool;
   END_VAR
   VAR_TEMP
      Stamp : DTL;
      ResultCode : Int;
   END_VAR
BEGIN

   #FRK_State := #Ok;
   IF #Idx < 1 OR #Idx > 12 OR LEN(#Key) = 0 OR LEN(#Key) > 120 THEN
       RETURN;
   END_IF;
   IF #Idx > #Count THEN
       #Count := #Idx;
   END_IF;
   IF #Flags[#Idx].Value <> #Ok OR #Flags[#Idx].Key <> #Key OR #Flags[#Idx].Stale THEN
       #Flags[#Idx].Since := LDT#1970-01-01-00:00:00.000000000;
       #ResultCode := RD_SYS_T(OUT => #Stamp);
       IF #ResultCode = 0 THEN
           #Flags[#Idx].Since := DTL_TO_LDT(#Stamp);
       END_IF;
   END_IF;
   #Flags[#Idx].Key := #Key;
   #Flags[#Idx].Value := #Ok;
   #Flags[#Idx].Stale := FALSE;
   #Touched[#Idx] := TRUE;
END_FUNCTION

FUNCTION "FRK_StateSweep" : Void   // FC20, SCL
{ S7_Optimized_Access := 'TRUE' }
VERSION : 0.1
// Core 3.12: derived facts; owning frame resolves freshness every scan.
// stored: AutoNumber true, IsIECCheckEnabled false, SetENOAutomatically false, UDAEnableTagReadback false
   VAR_INPUT
      Startup : Bool;
   END_VAR
   VAR_IN_OUT
      Flags : Array[1..12] of "ST_StateFlag";
      Count : Int;
      Touched : Array[1..12] of Bool;
   END_VAR
   VAR_TEMP
      Index : Int;
   END_VAR
BEGIN

   IF #Count < 0 OR #Count > 12 THEN
       #Count := 0;
   END_IF;
   FOR #Index := 1 TO #Count DO
       IF #Startup OR NOT #Touched[#Index] THEN
           #Flags[#Index].Value := FALSE;
           #Flags[#Index].Stale := TRUE;
       END_IF;
       #Touched[#Index] := FALSE;
   END_FOR;
END_FUNCTION

FUNCTION "FRK_SyncRegistry" : Void   // FC2, SCL
{ S7_Optimized_Access := 'TRUE' }
VERSION : 0.1
// stored: AutoNumber true, IsIECCheckEnabled false, SetENOAutomatically false, UDAEnableTagReadback false
   VAR_INPUT
      Index : DInt;
      Status : "ST_ModuleStatus";
   END_VAR
BEGIN

   // Nested checks precede array access; do not depend on short-circuit AND.
   IF #Index < 1 OR #Index > "FRK_Registry".Count OR #Index > 4 THEN
       "FRK_Registry".Fault := TRUE;
       RETURN;
   END_IF;
   IF NOT "FRK_Registry".Rows[#Index].Valid THEN
       "FRK_Registry".Fault := TRUE;
       RETURN;
   END_IF;
   "FRK_Registry".Rows[#Index].Exec := #Status.State;
   "FRK_Registry".Rows[#Index].ReasonCode := #Status.Diagnostic.ReasonCode;
   "FRK_Registry".Rows[#Index].Severity := #Status.Diagnostic.Severity;
END_FUNCTION

FUNCTION "FRK_UnitCascade" : Void   // FC84, SCL
{ S7_Optimized_Access := 'TRUE' }
VERSION : 0.1
// stored: AutoNumber true, IsIECCheckEnabled false, SetENOAutomatically false, UDAEnableTagReadback false
   VAR_INPUT
      ParentUnit : "FRK_Unit";
      Supported : Array[0..6] of Bool;
   END_VAR
   VAR_IN_OUT
      Core : "FRK_Core";
      Unit : "FRK_Unit";
      Status : "ST_ModuleStatus";
      Policy : Array[0..6] of "ST_ModePolicy";
      Access : "FRK_Access";
      AlarmLog : "FRK_AlarmLog";
   END_VAR
   VAR_TEMP
      Request : "ST_HmiRequest";
   END_VAR
BEGIN

   IF NOT #ParentUnit.CascadePending THEN
       RETURN;
   END_IF;
   IF #ParentUnit.CascadeKind = 6 OR #ParentUnit.CascadeKind = 9 THEN
       #Unit.FollowStart := FALSE;
       #Request.Kind := #ParentUnit.CascadeKind;
       "FRK_UnitOperation"(Core := #Core,
                           Unit := #Unit,
                           Status := #Status,
                           Policy := #Policy,
                           Access := #Access,
                           Supported := #Supported,
                           Request := #Request,
                           Response := "FRK_UnitScratch".Response,
                           Trusted := TRUE);
       RETURN;
   END_IF;
   #Request.Kind := 3;
   #Request.IntValue := #ParentUnit.CascadeMode;
   "FRK_UnitOperation"(Core := #Core,
                       Unit := #Unit,
                       Status := #Status,
                       Policy := #Policy,
                       Access := #Access,
                       Supported := #Supported,
                       Request := #Request,
                       Response := "FRK_UnitScratch".Response,
                       Trusted := TRUE);
   IF NOT "FRK_UnitScratch".Response.Accepted THEN
       #Unit.FollowStart := FALSE;
       #Request.Kind := 6;
       "FRK_UnitOperation"(Core := #Core,
                           Unit := #Unit,
                           Status := #Status,
                           Policy := #Policy,
                           Access := #Access,
                           Supported := #Supported,
                           Request := #Request,
                           Response := "FRK_UnitScratch".Response,
                           Trusted := TRUE);
       // Core names this event but has no assigned E_Reason ordinal yet.
       "FRK_AlarmMessage"(AlarmLog := #AlarmLog,
                          Reason := 2008,
                          Description := WSTRING#'std.event.childModeUnsupported',
                          SourcePath := STRING_TO_WSTRING(#Status.Name));
   ELSE
       #Unit.FollowStart := #ParentUnit.CascadeKind = 5;
   END_IF;
END_FUNCTION

FUNCTION "FRK_UnitConsume" : Void   // FC72, SCL
{ S7_Optimized_Access := 'TRUE' }
VERSION : 0.1
// stored: AutoNumber true, IsIECCheckEnabled false, SetENOAutomatically false, UDAEnableTagReadback false
   VAR_INPUT
      Supported : Array[0..6] of Bool;
   END_VAR
   VAR_IN_OUT
      Core : "FRK_Core";
      Unit : "FRK_Unit";
      Status : "ST_ModuleStatus";
      Policy : Array[0..6] of "ST_ModePolicy";
      Access : "FRK_Access";
      Response : "ST_HmiResponse";
   END_VAR
BEGIN

   IF NOT #Unit.RequestPending THEN
       RETURN;
   END_IF;
   // The generated typed ownership walk serves the static manifest after children.
   IF #Unit.Request.Kind = 23 THEN
       #Unit.Request.Secret := '';
       RETURN;
   END_IF;
   "FRK_UnitOperation"(Core := #Core,
                       Unit := #Unit,
                       Status := #Status,
                       Policy := #Policy,
                       Access := #Access,
                       Supported := #Supported,
                       Request := #Unit.Request,
                       Response := #Response,
                       Trusted := FALSE);
   #Unit.Request.Secret := '';
END_FUNCTION

FUNCTION "FRK_UnitFinish" : Void   // FC77, SCL
{ S7_Optimized_Access := 'TRUE' }
VERSION : 0.1
// stored: AutoNumber true, IsIECCheckEnabled false, SetENOAutomatically false, UDAEnableTagReadback false
   VAR_IN_OUT
      Core : "FRK_Core";
      Unit : "FRK_Unit";
      Response : "ST_HmiResponse";
      Status : "ST_ModuleStatus";
      Part : "ST_PartContext";
      AlarmLog : "FRK_AlarmLog";
      History : Array[1..16] of "ST_Diagnostic";
      Head : Int;
   END_VAR
BEGIN

   IF #Core.Exec = 3 THEN
       IF NOT #Unit.EvReset THEN
           #Unit.FaultLatched := TRUE;
       END_IF;
       IF NOT #Unit.PrevError THEN
           IF #Head < 0 OR #Head >= 16 THEN
               #Head := 0;
           END_IF;
           #Head := #Head + 1;
           #History[#Head] := #Status.Diagnostic;
           "FRK_PartAborted"(Core := #Core,
                             Unit := #Unit,
                             Status := #Status,
                             Part := #Part,
                             AlarmLog := #AlarmLog);
       END_IF;
   END_IF;
   #Unit.PrevError := #Core.Exec = 3;
   IF #Core.Exec = 2 OR #Core.Exec = 4 THEN
       #Unit.RunReq := FALSE;
   END_IF;
   IF #Unit.Clearing AND #Core.Exec = 0 THEN
       IF "FRK_DescendantsReady"(OwnerIndex := #Core.RegIndex) THEN
           #Unit.Clearing := FALSE;
       END_IF;
   END_IF;
   #Unit.AbortReq := FALSE;
   #Unit.ReleaseChildren := FALSE;
   #Unit.EvReset := FALSE;
   IF #Unit.RequestPending THEN
       #Response.AckSequence := #Unit.SeenSequence;
       #Unit.RequestPending := FALSE;
   END_IF;
END_FUNCTION

FUNCTION "FRK_UnitFollow" : Void   // FC85, SCL
{ S7_Optimized_Access := 'TRUE' }
VERSION : 0.1
// stored: AutoNumber true, IsIECCheckEnabled false, SetENOAutomatically false, UDAEnableTagReadback false
   VAR_INPUT
      Supported : Array[0..6] of Bool;
   END_VAR
   VAR_IN_OUT
      Core : "FRK_Core";
      Unit : "FRK_Unit";
      Status : "ST_ModuleStatus";
      Policy : Array[0..6] of "ST_ModePolicy";
      Access : "FRK_Access";
   END_VAR
   VAR_TEMP
      Request : "ST_HmiRequest";
   END_VAR
BEGIN

   IF #Unit.FollowStart AND NOT #Unit.ModePending AND NOT #Unit.Clearing THEN
       #Unit.FollowStart := FALSE;
       #Request.Kind := 5;
       "FRK_UnitOperation"(Core := #Core,
                           Unit := #Unit,
                           Status := #Status,
                           Policy := #Policy,
                           Access := #Access,
                           Supported := #Supported,
                           Request := #Request,
                           Response := "FRK_UnitScratch".Response,
                           Trusted := TRUE);
   END_IF;
END_FUNCTION

FUNCTION "FRK_UnitMailbox" : Void   // FC71, SCL
{ S7_Optimized_Access := 'TRUE' }
VERSION : 0.1
// stored: AutoNumber true, IsIECCheckEnabled false, SetENOAutomatically false, UDAEnableTagReadback false
   VAR_INPUT
      Supported : Array[0..6] of Bool;
   END_VAR
   VAR_IN_OUT
      Core : "FRK_Core";
      Unit : "FRK_Unit";
      Status : "ST_ModuleStatus";
      Policy : Array[0..6] of "ST_ModePolicy";
      Access : "FRK_Access";
      Request : "ST_HmiRequest";
      Response : "ST_HmiResponse";
   END_VAR
   VAR_TEMP
      SequenceBefore : UDInt;
   END_VAR
BEGIN

   #SequenceBefore := #Request.Sequence;
   IF #SequenceBefore = 0 OR #SequenceBefore = #Unit.SeenSequence THEN
       RETURN;
   END_IF;
   #Unit.Request := #Request;
   IF #Request.Sequence <> #SequenceBefore THEN
       #Unit.Request.Secret := '';
       RETURN;
   END_IF;
   #Request.Secret := '';
   #Unit.RequestUser := #Access.CurrentUser;
   #Unit.SeenSequence := #SequenceBefore;
   #Unit.RequestPending := TRUE;
END_FUNCTION

FUNCTION "FRK_UnitMode" : Void   // FC73, SCL
{ S7_Optimized_Access := 'TRUE' }
VERSION : 0.1
// stored: AutoNumber true, IsIECCheckEnabled false, SetENOAutomatically false, UDAEnableTagReadback false
   VAR_IN_OUT
      Core : "FRK_Core";
      Unit : "FRK_Unit";
   END_VAR
BEGIN

   IF #Unit.ModePending THEN
       IF #Core.Exec = 1 THEN
           #Core.EvModeExit := TRUE;
           #Core.HookResult := 0;
       ELSIF #Core.Exec = 0 AND NOT #Unit.Clearing THEN
           #Unit.Mode := #Unit.RequestedMode;
           #Unit.ModePending := FALSE;
           #Unit.ExitFirst := FALSE;
           #Core.EvModeChanged := TRUE;
       ELSE
           #Unit.RunReq := FALSE;
       END_IF;
   END_IF;
END_FUNCTION

FUNCTION "FRK_UnitModeResolve" : Void   // FC74, SCL
{ S7_Optimized_Access := 'TRUE' }
VERSION : 0.1
// stored: AutoNumber true, IsIECCheckEnabled false, SetENOAutomatically false, UDAEnableTagReadback false
   VAR_INPUT
      Policy : Array[0..6] of "ST_ModePolicy";
      Timeout : Time;
   END_VAR
   VAR_IN_OUT
      Core : "FRK_Core";
      Unit : "FRK_Unit";
      Status : "ST_ModuleStatus";
   END_VAR
BEGIN

   IF #Unit.ModePending THEN
       IF #Timeout <= T#0ms OR "FRK_Elapsed"(NewMs := "FRK_Clock".NowMs, OldMs := #Unit.ModeSince) >= DINT_TO_UDINT(TIME_TO_DINT(#Timeout)) THEN
           "FRK_Fault"(Core := #Core,
                       Status := #Status,
                       ReasonCode := 2001,
                       Description := WSTRING#'std.error.hmiRequestRejected');
           #Unit.ModePending := FALSE;
           #Unit.FollowStart := FALSE;
           #Unit.ReleaseChildren := TRUE;
           #Unit.Clearing := TRUE;
       ELSIF #Core.EvModeExit THEN
           #Unit.ExitFirst := FALSE;
           IF #Policy[#Unit.Mode].Style = 0 THEN
               #Unit.StopReq := TRUE;
           ELSIF #Core.HookResult <= 0 THEN
               #Unit.AbortReq := TRUE;
               #Unit.ReleaseChildren := TRUE;
               #Unit.Clearing := TRUE;
           END_IF;
       END_IF;
   END_IF;
END_FUNCTION

FUNCTION "FRK_UnitOperation" : Void   // FC70, SCL
{ S7_Optimized_Access := 'TRUE' }
VERSION : 0.1
// stored: AutoNumber true, IsIECCheckEnabled false, SetENOAutomatically false, UDAEnableTagReadback false
   VAR_INPUT
      Supported : Array[0..6] of Bool;
      Request : "ST_HmiRequest";
      Trusted : Bool;
   END_VAR
   VAR_IN_OUT
      Core : "FRK_Core";
      Unit : "FRK_Unit";
      Status : "ST_ModuleStatus";
      Policy : Array[0..6] of "ST_ModePolicy";
      Access : "FRK_Access";
      Response : "ST_HmiResponse";
   END_VAR
   VAR_TEMP
      Gate : DInt;
      Desired : DInt;
      Query : Bool;
      Level : DInt;
      DecisionAccepted : Bool;
   END_VAR
BEGIN

   #Response.Accepted := FALSE;
   #Response.Diagnostic := WSTRING#'';
   #Response.Report.Count := 0;
   #Response.Report.Released := TRUE;
   #Gate := -1;
   #Desired := -1;
   #Query := FALSE;
   CASE #Request.Kind OF
       5:
           #Gate := 5;
           #Desired := 0;
       6:
           #Gate := 5;
           #Desired := 1;
       3:
           #Gate := 4;
           #Desired := #Request.IntValue;
           IF #Desired = -1 THEN
               #Desired := -2;
           END_IF;
       9:
           #Gate := 7;
       10:
           #Gate := 5;
       11:
           #Gate := 2;
       24, 25:
           #Gate := 8;
       15:
           #Gate := 5;
           #Desired := 0;
           #Query := TRUE;
       16:
           #Gate := 2;
           #Query := TRUE;
       17:
           #Gate := #Request.IntValue;
           #Desired := -1;
           #Query := TRUE;
       ELSE
           #Gate := -1;
   END_CASE;
   IF #Gate <> -1 OR #Request.Kind = 17 THEN
       "FRK_UnitRelease"(Core := #Core,
                         Unit := #Unit,
                         Status := #Status,
                         Policy := #Policy,
                         Access := #Access,
                         Supported := #Supported,
                         Report := #Response.Report,
                         Gate := #Gate,
                         Desired := #Desired,
                         Trusted := #Trusted);
       IF #Query THEN
           #Response.Accepted := TRUE;
       ELSIF #Response.Report.Released THEN
           CASE #Request.Kind OF
               10:
                   #DecisionAccepted := "FRK_DecisionSubmit"(Owner := #Core.RegIndex,
                                                             OwnerPath := STRING_TO_WSTRING(#Status.Name),
                                                             Option := #Request.IntValue,
                                                             Busy := #Core.Exec = 1,
                                                             Permit := #Unit.Permit,
                                                             Report := #Response.Report);
                   #Response.Accepted := #DecisionAccepted;
               5:
                   #Unit.StopReq := FALSE;
                   #Unit.RunReq := TRUE;
                   #Response.Accepted := TRUE;
               6:
                   #Unit.StopReq := #Core.Exec = 1;
                   IF NOT #Unit.StopReq THEN
                       #Unit.RunReq := FALSE;
                   END_IF;
                   #Unit.FollowStart := FALSE;
                   #Response.Accepted := TRUE;
               3:
                   IF #Desired <> #Unit.Mode THEN
                       #Unit.ExitFirst := TRUE;
                       #Unit.ModeSince := "FRK_Clock".NowMs;
                       #Unit.RequestedMode := #Desired;
                       #Unit.ModePending := TRUE;
                       IF #Unit.Mode = 1 THEN
                           #Unit.ReleaseChildren := TRUE;
                           #Unit.Clearing := TRUE;
                       END_IF;
                   END_IF;
                   #Response.Accepted := TRUE;
               9:
                   #Unit.EvReset := TRUE;
                   #Unit.ModePending := FALSE;
                   #Unit.ExitFirst := FALSE;
                   #Unit.RunReq := FALSE;
                   #Unit.AbortReq := #Core.Exec = 1;
                   #Unit.StopReq := FALSE;
                   #Unit.FollowStart := FALSE;
                   #Unit.ReleaseChildren := TRUE;
                   #Unit.Clearing := TRUE;
                   #Unit.FaultLatched := FALSE;
                   IF #Core.Exec = 3 THEN
                       #Core.Armed := TRUE;
                   END_IF;
                   #Response.Accepted := TRUE;
               24:
                   #Level := -1;
                   IF #Request.TextValue = WSTRING#'0' THEN
                       #Level := 0;
                   ELSIF #Request.TextValue = WSTRING#'1' THEN
                       #Level := 1;
                   ELSIF #Request.TextValue = WSTRING#'2' THEN
                       #Level := 2;
                   ELSIF #Request.TextValue = WSTRING#'3' THEN
                       #Level := 3;
                   ELSIF #Request.TextValue = WSTRING#'4' THEN
                       #Level := 4;
                   END_IF;
                   IF #Request.IntValue >= 0 AND #Request.IntValue <= 11 AND #Level >= 0 THEN
                       IF #Request.IntValue <> 8 OR #Level <= #Access.CurrentLevel THEN
                           #Access.Policy.Required[#Request.IntValue] := #Level;
                           #Response.Accepted := TRUE;
                       END_IF;
                   END_IF;
               25:
                   IF #Request.DurationMs <= 604800000 THEN
                       #Access.Policy.SessionTimeout := DINT_TO_TIME(UDINT_TO_DINT(#Request.DurationMs));
                       #Response.Accepted := TRUE;
                   END_IF;
               ELSE
                   // Manual acceptance is resolved by the generated typed route.
                   #Response.Accepted := FALSE;
           END_CASE;
       END_IF;
   ELSE
       CASE #Request.Kind OF
           1:
               "FRK_AccessLogin"(Access := #Access,
                                 User := #Request.User,
                                 Secret := #Request.Secret,
                                 Sequence := #Request.Sequence);
               // Consumption is acknowledged now; correlated result is asynchronous.
               #Response.Accepted := TRUE;
           2:
               "FRK_AccessLogout"(Access := #Access);
               #Response.Accepted := TRUE;
           ELSE
               #Response.Diagnostic := WSTRING#'std.error.unsupportedHmiRequest';
       END_CASE;
   END_IF;
   IF #Response.Accepted AND NOT #Query THEN
       IF #Request.Kind = 5 OR #Request.Kind = 6 OR #Request.Kind = 3 OR #Request.Kind = 9 THEN
           #Unit.CascadePending := TRUE;
           #Unit.CascadeKind := #Request.Kind;
           #Unit.CascadeMode := #Unit.Mode;
           IF #Request.Kind = 3 THEN
               #Unit.CascadeMode := #Desired;
           END_IF;
       END_IF;
   END_IF;
   IF NOT #Response.Accepted AND #Request.Kind <> 11 THEN
       IF #Response.Diagnostic = WSTRING#'' THEN
           #Response.Diagnostic := WSTRING#'std.error.hmiRequestRejected';
       END_IF;
       IF #Response.Report.Released THEN
           "FRK_ReleaseReason"(Report := #Response.Report,
                               Description := #Response.Diagnostic,
                               Reason := 2002,
                               Path := STRING_TO_WSTRING(#Status.Name),
                               Kind := 4);
       END_IF;
   END_IF;
END_FUNCTION

FUNCTION "FRK_UnitPrepare" : Void   // FC61, SCL
{ S7_Optimized_Access := 'TRUE' }
VERSION : 0.1
// Shared Unit services v0.1: operation authority, mailbox, modes and local carrier.
// stored: AutoNumber true, IsIECCheckEnabled false, SetENOAutomatically false, UDAEnableTagReadback false
   VAR_INPUT
      Startup : Bool;
      InitialMode : DInt;
   END_VAR
   VAR_IN_OUT
      Core : "FRK_Core";
      Unit : "FRK_Unit";
      Policy : Array[0..6] of "ST_ModePolicy";
      Request : "ST_HmiRequest";
      Response : "ST_HmiResponse";
   END_VAR
   VAR_TEMP
      Index : DInt;
   END_VAR
BEGIN

   #Core.EvModeExit := FALSE;
   #Core.EvModeChanged := FALSE;
   IF NOT #Unit.Initialized THEN
       #Unit.Initialized := TRUE;
       #Unit.Permit := TRUE;
       FOR #Index := 0 TO 7 - 1 DO
           #Policy[#Index].Shield := 1;
           #Policy[#Index].Style := 1;
       END_FOR;
       #Policy[0].Style := 0;
       #Policy[2].Shield := 0;
       #Policy[1].Shield := 0;
       #Policy[3].Shield := 2;
       #Policy[4].Shield := 2;
       #Unit.Mode := #InitialMode;
   END_IF;
   IF #Startup THEN
       #Unit.EvReset := FALSE;
       #Unit.Mode := #InitialMode;
       #Unit.RunReq := FALSE;
       #Unit.AbortReq := #Core.Exec = 1;
       #Unit.StopReq := FALSE;
       #Unit.ModePending := FALSE;
       #Unit.FollowStart := FALSE;
       #Unit.CascadePending := FALSE;
       #Unit.ReleaseChildren := TRUE;
       #Unit.Clearing := TRUE;
       // Consume the restart boundary without executing a transported request.
       #Unit.SeenSequence := #Request.Sequence;
       #Unit.RequestPending := FALSE;
       #Request.Secret := '';
       #Response.Accepted := FALSE;
       #Response.Diagnostic := WSTRING#'std.error.hmiRequestRejected';
       #Response.AckSequence := #Unit.SeenSequence;
   END_IF;
   IF #Core.ReleasePending THEN
       #Unit.FollowStart := FALSE;
       // An incoming parent mode/reset operation is already queued for this scan.
       // Preserve its cascade while cancelling the old command.
       #Unit.RunReq := FALSE;
       #Unit.AbortReq := TRUE;
       #Unit.ReleaseChildren := TRUE;
       #Unit.Clearing := TRUE;
   END_IF;
END_FUNCTION

